(* IEC 61131-3 sources: RootPLC/conformance/cases/blocks, 22 files *)

(* ---- ok_rb_round4.st ---- *)
(* spec: [blocks.fault] [blocks.testable]
   expect: ok
   libraries: RootBlocks *)
(* Test suites of RB_SetpointProfile (F06.PROFILE), RB_Homing (F05.HOMING),
   RB_DataLog (F11.LOG), RB_ScaleOut (F01.SCALE.OUT) and RB_Drum
   (F05.DRUM). Every call passes the inputs that matter: block inputs keep
   their last value. *)
FUNCTION_BLOCK FB_Profile2
VAR_OUTPUT
    tg : ARRAY[1..8] OF REAL;
    rt : ARRAY[1..8] OF TIME;
    st : ARRAY[1..8] OF TIME;
END_VAR
tg[1] := 100.0; rt[1] := T#10s; st[1] := T#5s;
tg[2] := 50.0;  rt[2] := T#5s;  st[2] := T#2s;
END_FUNCTION_BLOCK

TEST profile_ramps_and_soaks
VAR p : RB_SetpointProfile; d : FB_Profile2; END_VAR
d();
p(PV := 20.0, Count := 2, Targets := d.tg, RampTimes := d.rt, SoakTimes := d.st);
ASSERT_FALSE(p.Busy);
ASSERT_EQ(0, p.Segment);
ADVANCE(T#1s);
p(Start := TRUE);
ASSERT_TRUE(p.Busy);
ASSERT_EQ(1, p.Segment);
ASSERT_TRUE(ABS(p.SP - 20.0) < 0.001);
ADVANCE(T#5s);
p(Start := FALSE);
ASSERT_TRUE(ABS(p.SP - 60.0) < 0.01);
ASSERT_FALSE(p.Soaking);
ADVANCE(T#5s);
p();
ASSERT_TRUE(ABS(p.SP - 100.0) < 0.001);
ASSERT_TRUE(p.Soaking);
ADVANCE(T#4900ms);
p();
ASSERT_EQ(1, p.Segment);
ADVANCE(T#100ms);
p();
ASSERT_EQ(2, p.Segment);
ASSERT_FALSE(p.Soaking);
ADVANCE(T#2500ms);
p();
ASSERT_TRUE(ABS(p.SP - 75.0) < 0.01);
ADVANCE(T#2500ms);
p();
ASSERT_TRUE(ABS(p.SP - 50.0) < 0.001);
ADVANCE(T#2s);
p();
ASSERT_TRUE(p.Done);
ASSERT_FALSE(p.Busy);
ASSERT_EQ(0, p.Segment);
ASSERT_TRUE(ABS(p.SP - 50.0) < 0.001);
(* a new start clears Done *)
p(Start := TRUE, PV := 30.0);
ASSERT_FALSE(p.Done);
ASSERT_TRUE(ABS(p.SP - 30.0) < 0.001);
END_TEST

TEST profile_hold_guarantee_and_abort
VAR p : RB_SetpointProfile; d : FB_Profile2; END_VAR
d();
p(PV := 20.0, Count := 1, Targets := d.tg, RampTimes := d.rt, SoakTimes := d.st, Start := TRUE);
ADVANCE(T#5s);
p(Start := FALSE);
ASSERT_TRUE(ABS(p.SP - 60.0) < 0.01);
ADVANCE(T#10s);
p(Hold := TRUE);
ASSERT_TRUE(ABS(p.SP - 60.0) < 0.01);
p(Hold := FALSE);
ADVANCE(T#5s);
p(Band := 2.0);
ASSERT_TRUE(p.Soaking);
(* guaranteed soak: PV far from SP, the soak waits *)
ADVANCE(T#10s);
p(PV := 90.0);
ASSERT_TRUE(p.Soaking);
ASSERT_EQ(1, p.Segment);
ADVANCE(T#1s);
p(PV := 98.0);
(* each call counts the time since the previous one *)
ADVANCE(T#3s);
p(PV := 98.0);
ASSERT_TRUE(p.Busy);
ADVANCE(T#1s);
p(PV := 98.0);
ASSERT_TRUE(p.Done);
(* abort while soaking *)
p(Start := TRUE, PV := 100.0);
ASSERT_TRUE(p.Busy);
ADVANCE(T#10s);
p(Start := FALSE);
ASSERT_TRUE(p.Soaking);
p(Abort := TRUE);
ASSERT_FALSE(p.Soaking);
ASSERT_FALSE(p.Busy);
ASSERT_EQ(0, p.Segment);
ASSERT_FALSE(p.Done);
ADVANCE(T#20s);
p(Abort := FALSE);
ASSERT_FALSE(p.Busy);
END_TEST

TEST profile_zero_times_and_count
VAR p : RB_SetpointProfile; tg : ARRAY[1..8] OF REAL; rt, st : ARRAY[1..8] OF TIME; END_VAR
tg[1] := 70.0;
p(PV := 10.0, Count := 0, Targets := tg, RampTimes := rt, SoakTimes := st, Start := TRUE);
ASSERT_TRUE(p.Error);
ASSERT_EQ(UDINT#1, p.ErrorID);
ASSERT_FALSE(p.Busy);
p(Start := FALSE, Count := 9);
p(Start := TRUE);
ASSERT_TRUE(p.Error);
p(Start := FALSE, Count := 8);
p(Start := TRUE);
ASSERT_FALSE(p.Error);
ASSERT_EQ(UDINT#0, p.ErrorID);
(* T#0s ramp and soak: a step to the target, one segment per call *)
p(Start := FALSE);
ASSERT_TRUE(ABS(p.SP - 70.0) < 0.001);
p();
ASSERT_EQ(2, p.Segment);
p(Count := 1);
p();
ASSERT_TRUE(p.Done);
(* a start with a bad count while running ends the program *)
p(Count := 8);
p(Start := TRUE);
p(Start := FALSE);
p();
ASSERT_EQ(2, p.Segment);
p(Count := 0);
p(Start := TRUE);
ASSERT_EQ(0, p.Segment);
ASSERT_FALSE(p.Busy);
END_TEST

TEST homing_seeks_and_backs_off
VAR h : RB_Homing; END_VAR
h();
ASSERT_FALSE(h.Busy OR h.Homed);
h(Start := TRUE);
ASSERT_TRUE(h.MoveToHome);
ASSERT_FALSE(h.MoveAway OR h.Slow);
ASSERT_TRUE(h.Busy);
ADVANCE(T#20s);
h(Start := FALSE, HomeSwitch := TRUE);
ASSERT_FALSE(h.MoveToHome);
ASSERT_TRUE(h.MoveAway AND h.Slow);
(* each phase has its own Timeout *)
ADVANCE(T#20s);
h();
ASSERT_FALSE(h.Error);
h(HomeSwitch := FALSE);
ASSERT_TRUE(h.Homed);
ASSERT_FALSE(h.Busy OR h.MoveAway OR h.MoveToHome);
(* starting on the switch: straight to backing off; Homed clears *)
h(Start := TRUE, HomeSwitch := TRUE);
ASSERT_FALSE(h.Homed);
ASSERT_TRUE(h.MoveAway);
h(Start := FALSE, HomeSwitch := FALSE);
ASSERT_TRUE(h.Homed);
(* a new start while seeking restarts the timing *)
h(Start := TRUE, Timeout := T#2s);
ADVANCE(T#1500ms);
h(Start := FALSE);
h(Start := TRUE);
ADVANCE(T#1500ms);
h(Start := FALSE);
ASSERT_FALSE(h.Error);
ASSERT_TRUE(h.MoveToHome);
h(Timeout := T#30s);
(* abort *)
h(Start := TRUE);
ASSERT_TRUE(h.MoveToHome);
h(Start := FALSE, Abort := TRUE);
ASSERT_FALSE(h.Busy OR h.MoveToHome OR h.Homed);
h(Start := TRUE);
ASSERT_FALSE(h.Busy);
END_TEST

TEST homing_timeouts
VAR h : RB_Homing; END_VAR
h(Start := TRUE, Timeout := T#2s);
ADVANCE(T#1900ms);
h();
ASSERT_FALSE(h.Error);
ADVANCE(T#100ms);
h();
ASSERT_TRUE(h.Error);
ASSERT_EQ(UDINT#1, h.ErrorID);
ASSERT_FALSE(h.MoveToHome OR h.Busy);
(* no start while the fault lasts *)
h(Start := FALSE);
h(Start := TRUE);
ASSERT_FALSE(h.Busy);
h(Start := FALSE, Reset := TRUE);
ASSERT_FALSE(h.Error);
ASSERT_EQ(UDINT#0, h.ErrorID);
h(Reset := FALSE, Start := TRUE);
ASSERT_TRUE(h.MoveToHome);
h(Start := FALSE, HomeSwitch := TRUE);
ADVANCE(T#2s);
h();
ASSERT_TRUE(h.Error);
ASSERT_EQ(UDINT#2, h.ErrorID);
ASSERT_FALSE(h.MoveAway OR h.Slow);
ASSERT_FALSE(h.Homed);
END_TEST

TEST data_log_ring_and_statistics
VAR l : RB_DataLog; i : INT; END_VAR
l(Value := 0.0, Enable := FALSE);
ASSERT_EQ(0, l.Count);
ASSERT_EQ(0, l.Newest);
l(Value := 5.0, Enable := TRUE);
ASSERT_EQ(1, l.Count);
ASSERT_EQ(1, l.Newest);
ASSERT_TRUE(ABS(l.Minimum - 5.0) < 0.001 AND ABS(l.Maximum - 5.0) < 0.001 AND ABS(l.Average - 5.0) < 0.001);
ADVANCE(T#500ms);
l(Value := 9.0);
ASSERT_EQ(1, l.Count);
ADVANCE(T#500ms);
l(Value := 1.0);
ASSERT_EQ(2, l.Count);
ASSERT_TRUE(ABS(l.Samples[2] - 1.0) < 0.001);
ASSERT_TRUE(ABS(l.Minimum - 1.0) < 0.001);
ASSERT_TRUE(ABS(l.Maximum - 5.0) < 0.001);
ASSERT_TRUE(ABS(l.Average - 3.0) < 0.001);
(* fill and wrap: 70 samples in all *)
FOR i := 3 TO 70 DO
    ADVANCE(T#1s);
    l(Value := INT_TO_REAL(i));
END_FOR;
ASSERT_EQ(64, l.Count);
ASSERT_EQ(6, l.Newest);
ASSERT_TRUE(ABS(l.Samples[6] - 70.0) < 0.001);
ASSERT_TRUE(ABS(l.Minimum - 7.0) < 0.001);
ASSERT_TRUE(ABS(l.Maximum - 70.0) < 0.001);
ASSERT_TRUE(ABS(l.Average - 38.5) < 0.001);
(* the next sample comes one Interval later, not before *)
ADVANCE(T#500ms);
l(Value := 71.0);
ASSERT_EQ(6, l.Newest);
ADVANCE(T#500ms);
l(Value := 71.0);
ASSERT_EQ(7, l.Newest);
(* paused, then cleared *)
ADVANCE(T#5s);
l(Value := 99.0, Enable := FALSE);
ASSERT_TRUE(ABS(l.Maximum - 71.0) < 0.001);
l(Clear := TRUE);
ASSERT_EQ(0, l.Count);
ASSERT_TRUE(ABS(l.Average) < 0.001 AND ABS(l.Maximum) < 0.001 AND ABS(l.Minimum) < 0.001);
l(Clear := FALSE, Enable := TRUE, Value := -4.0);
ASSERT_EQ(1, l.Newest);
ASSERT_TRUE(ABS(l.Minimum + 4.0) < 0.001 AND ABS(l.Maximum + 4.0) < 0.001);
END_TEST

TEST scale_out_to_an_output_word
VAR s : RB_ScaleOut; END_VAR
s(Value := 50.0);
ASSERT_EQ(13824, s.Raw);
ASSERT_FALSE(s.Limited OR s.Error);
s(Value := 100.0);
ASSERT_EQ(27648, s.Raw);
ASSERT_FALSE(s.Limited);
s(Value := 120.0);
ASSERT_EQ(27648, s.Raw);
ASSERT_TRUE(s.Limited);
s(Value := -5.0);
ASSERT_EQ(0, s.Raw);
ASSERT_TRUE(s.Limited);
s(Value := 0.5);
ASSERT_EQ(138, s.Raw);
s(Value := 0.0);
ASSERT_EQ(0, s.Raw);
ASSERT_FALSE(s.Limited);
(* the fail value on a fault *)
s(Value := 50.0, Fault := TRUE, FailValue := 25.0);
ASSERT_EQ(6912, s.Raw);
s(Fault := FALSE);
ASSERT_EQ(13824, s.Raw);
(* a reversed range and a live-zero raw range *)
s(Value := 25.0, EngMin := 100.0, EngMax := 0.0);
ASSERT_EQ(20736, s.Raw);
s(Value := 50.0, EngMin := 0.0, EngMax := 100.0, RawMin := 5530.0);
ASSERT_EQ(16589, s.Raw);
s(EngMax := 0.0);
ASSERT_TRUE(s.Error);
ASSERT_EQ(UDINT#1, s.ErrorID);
ASSERT_EQ(5530, s.Raw);
ASSERT_FALSE(s.Limited);
s(EngMax := 200.0);
ASSERT_FALSE(s.Error);
ASSERT_EQ(UDINT#0, s.ErrorID);
END_TEST

TEST drum_steps_by_time_and_event
VAR d : RB_Drum; p : ARRAY[1..16] OF WORD; t : ARRAY[1..16] OF TIME; END_VAR
p[1] := WORD#16#0001; p[2] := WORD#16#0006; p[3] := WORD#16#0010;
t[1] := T#2s; t[2] := T#0s; t[3] := T#1s;
d(Patterns := p, Times := t, Count := 3);
ASSERT_EQ(1, d.StepNo);
ASSERT_EQ(WORD#16#0001, d.Out);
ADVANCE(T#5s);
d();
ASSERT_EQ(1, d.StepNo);
d(Run := TRUE);
ADVANCE(T#1900ms);
d();
ASSERT_EQ(1, d.StepNo);
ASSERT_EQ(T#1900ms, d.StepTime);
ADVANCE(T#100ms);
d();
ASSERT_EQ(2, d.StepNo);
ASSERT_EQ(WORD#16#0006, d.Out);
ASSERT_EQ(T#0s, d.StepTime);
(* T#0s: waits for Next *)
ADVANCE(T#10s);
d();
ASSERT_EQ(2, d.StepNo);
d(Next := TRUE);
ASSERT_EQ(3, d.StepNo);
d(Next := FALSE);
(* paused while Run is FALSE *)
ADVANCE(T#500ms);
d();
ADVANCE(T#100ms);
d(Run := FALSE);
ADVANCE(T#100ms);
d(Run := FALSE);
ADVANCE(T#100ms);
d(Run := TRUE);
ADVANCE(T#300ms);
d();
ASSERT_EQ(3, d.StepNo);
ADVANCE(T#100ms);
d();
ASSERT_EQ(1, d.StepNo);
END_TEST

TEST drum_one_shot_reset_and_count
VAR d : RB_Drum; p : ARRAY[1..16] OF WORD; t : ARRAY[1..16] OF TIME; END_VAR
p[1] := WORD#16#00F0; p[2] := WORD#16#0F00;
d(Patterns := p, Times := t, Count := 2, Cyclic := FALSE);
d(Next := TRUE);
ASSERT_EQ(2, d.StepNo);
d(Next := FALSE);
d(Next := TRUE);
ASSERT_TRUE(d.Done);
ASSERT_EQ(2, d.StepNo);
ASSERT_EQ(WORD#16#0F00, d.Out);
d(Next := FALSE);
d(Next := TRUE);
ASSERT_EQ(2, d.StepNo);
d(Next := FALSE, Reset := TRUE);
ASSERT_EQ(1, d.StepNo);
ASSERT_FALSE(d.Done);
d(Reset := FALSE, Count := 0);
ASSERT_TRUE(d.Error);
ASSERT_EQ(UDINT#1, d.ErrorID);
ASSERT_EQ(WORD#0, d.Out);
ASSERT_EQ(0, d.StepNo);
d(Count := 17);
ASSERT_TRUE(d.Error);
d(Count := 1);
ASSERT_FALSE(d.Error);
ASSERT_EQ(1, d.StepNo);
d(Count := 16);
ASSERT_FALSE(d.Error);
ASSERT_EQ(UDINT#0, d.ErrorID);
ASSERT_EQ(1, d.StepNo);
(* a smaller Count while beyond it: back to step 1 *)
d(Next := TRUE);
d(Next := FALSE);
d(Next := TRUE);
d(Next := FALSE);
ASSERT_EQ(3, d.StepNo);
d(Count := 2);
ASSERT_EQ(1, d.StepNo);
END_TEST

(* ---- ok_rb_sequence.st ---- *)
(* spec: [blocks.command] [blocks.fault] [blocks.testable]
   expect: ok
   libraries: RootBlocks *)
(* Test suites of RB_StepChain (F05.STEPS) and RB_Phase (F05.PHASE). *)

(* the pattern the card shows: the chain, then the actions per step *)
FUNCTION_BLOCK FillCycle
VAR_INPUT
    start  : BOOL;
    full   : BOOL;
    empty  : BOOL;
END_VAR
VAR_OUTPUT
    inlet  : BOOL;
    outlet : BOOL;
    fills  : INT;
END_VAR
VAR
    chain : RB_StepChain;
END_VAR
CASE chain.StepNo OF
1: chain(Start := start, Proceed := full, LastStep := 2, StepTimeout := T#5s);
2: chain(Start := start, Proceed := empty, LastStep := 2, StepTimeout := T#5s);
ELSE
    chain(Start := start, Proceed := FALSE, LastStep := 2, StepTimeout := T#5s);
END_CASE;
inlet := chain.StepNo = 1;
outlet := chain.StepNo = 2;
IF chain.FirstCall AND chain.StepNo = 1 THEN
    fills := fills + 1;
END_IF;
END_FUNCTION_BLOCK

TEST chain_runs_its_steps_in_order
VAR f : FillCycle; END_VAR
f(start := FALSE);
ASSERT_EQ(0, f.chain.StepNo);
ASSERT_FALSE(f.chain.Busy);
f(start := TRUE);
ASSERT_EQ(1, f.chain.StepNo);
ASSERT_TRUE(f.inlet);
ASSERT_TRUE(f.chain.FirstCall);
ASSERT_TRUE(f.chain.Busy);
ASSERT_EQ(1, f.fills);
f(start := TRUE);
ASSERT_FALSE(f.chain.FirstCall);
ASSERT_EQ(1, f.fills);
f(start := TRUE, full := TRUE);
ASSERT_EQ(2, f.chain.StepNo);
ASSERT_TRUE(f.chain.FirstCall);
ASSERT_TRUE(f.outlet);
f(start := TRUE, full := TRUE, empty := TRUE);
ASSERT_EQ(0, f.chain.StepNo);
ASSERT_TRUE(f.chain.Done);
ASSERT_FALSE(f.chain.Busy);
f(start := TRUE, full := TRUE, empty := TRUE);
ASSERT_FALSE(f.chain.Done);
ASSERT_EQ(0, f.chain.StepNo);
(* a new rising edge starts it again *)
f(start := FALSE);
f(start := TRUE);
ASSERT_EQ(1, f.chain.StepNo);
ASSERT_EQ(2, f.fills);
END_TEST

TEST chain_step_time_and_timeout
VAR c : RB_StepChain; END_VAR
c(Start := TRUE, LastStep := 3, StepTimeout := T#2s);
ADVANCE(T#1500ms);
c(Start := TRUE, LastStep := 3, StepTimeout := T#2s);
ASSERT_TRUE(c.StepTime = T#1500ms);
ASSERT_FALSE(c.Error);
ADVANCE(T#500ms);
c(Start := TRUE, LastStep := 3, StepTimeout := T#2s);
ASSERT_TRUE(c.Error);
ASSERT_EQ(UDINT#1, c.ErrorID);
ASSERT_EQ(1, c.StepNo);
(* the fault holds the chain: Proceed is ignored *)
c(Start := TRUE, Proceed := TRUE, LastStep := 3, StepTimeout := T#2s);
ASSERT_EQ(1, c.StepNo);
(* reset restarts the step timer *)
c(Start := TRUE, Proceed := FALSE, LastStep := 3, StepTimeout := T#2s, Reset := TRUE);
ASSERT_FALSE(c.Error);
ASSERT_EQ(UDINT#0, c.ErrorID);
ASSERT_TRUE(c.StepTime = T#0s);
ADVANCE(T#1s);
c(Start := TRUE, Proceed := TRUE, LastStep := 3, StepTimeout := T#2s, Reset := FALSE);
ASSERT_EQ(2, c.StepNo);
ASSERT_TRUE(c.StepTime = T#0s);
(* no timeout configured: no fault *)
ADVANCE(T#1h);
c(Start := TRUE, Proceed := FALSE, LastStep := 3, StepTimeout := T#0s);
ASSERT_FALSE(c.Error);
END_TEST

TEST chain_hold_pauses_and_abort_resets
VAR c : RB_StepChain; END_VAR
c(Start := TRUE, LastStep := 2, StepTimeout := T#2s);
ADVANCE(T#1s);
c(Start := TRUE, Hold := TRUE, Proceed := TRUE, LastStep := 2, StepTimeout := T#2s);
ASSERT_EQ(1, c.StepNo);
ASSERT_TRUE(c.Held);
ADVANCE(T#10s);
c(Start := TRUE, Hold := TRUE, Proceed := FALSE, LastStep := 2, StepTimeout := T#2s);
ASSERT_FALSE(c.Error);
ASSERT_TRUE(c.StepTime = T#0s);
c(Start := TRUE, Hold := FALSE, Proceed := FALSE, LastStep := 2, StepTimeout := T#2s);
ASSERT_FALSE(c.Held);
ASSERT_FALSE(c.Error);
c(Start := TRUE, Abort := TRUE, LastStep := 2, StepTimeout := T#2s);
ASSERT_EQ(0, c.StepNo);
ASSERT_TRUE(c.Aborted);
ASSERT_FALSE(c.Busy);
ASSERT_FALSE(c.Held);
c(Start := TRUE, Abort := TRUE, LastStep := 2, StepTimeout := T#2s);
ASSERT_FALSE(c.Aborted);
(* while Abort is TRUE the chain does not start *)
c(Start := FALSE, Abort := TRUE, LastStep := 2);
c(Start := TRUE, Abort := TRUE, LastStep := 2);
ASSERT_EQ(0, c.StepNo);
END_TEST

TEST chain_branches_with_next_step
VAR c : RB_StepChain; END_VAR
c(Start := TRUE, LastStep := 5);
c(Start := TRUE, Proceed := TRUE, NextStep := 4, LastStep := 5);
ASSERT_EQ(4, c.StepNo);
ASSERT_TRUE(c.FirstCall);
c(Start := TRUE, Proceed := TRUE, NextStep := 0, LastStep := 5);
ASSERT_EQ(5, c.StepNo);
(* a jump back from the last step keeps the chain running *)
c(Start := TRUE, Proceed := TRUE, NextStep := 2, LastStep := 5);
ASSERT_EQ(2, c.StepNo);
ASSERT_FALSE(c.Done);
(* an abort with an active timeout fault clears it *)
c(Start := TRUE, Proceed := FALSE, StepTimeout := T#1s, LastStep := 5);
ADVANCE(T#2s);
c(Start := TRUE, Proceed := FALSE, StepTimeout := T#1s, LastStep := 5);
ASSERT_TRUE(c.Error);
c(Start := TRUE, Abort := TRUE, LastStep := 5);
ASSERT_FALSE(c.Error);
ASSERT_EQ(UDINT#0, c.ErrorID);
END_TEST

TEST phase_runs_holds_and_completes
VAR p : RB_Phase; END_VAR
p();
ASSERT_TRUE(p.State = RB_PHASE_STATE#Idle);
p(Start := TRUE);
ASSERT_TRUE(p.State = RB_PHASE_STATE#Running);
ASSERT_TRUE(p.Running);
ASSERT_FALSE(p.Rejected);
p(Start := FALSE, Hold := TRUE);
ASSERT_TRUE(p.State = RB_PHASE_STATE#Held);
ASSERT_FALSE(p.Running);
p(Hold := FALSE, Finished := TRUE);
ASSERT_TRUE(p.State = RB_PHASE_STATE#Held);
p(Restart := TRUE, Finished := FALSE);
ASSERT_TRUE(p.State = RB_PHASE_STATE#Running);
p(Restart := FALSE, Finished := TRUE);
ASSERT_TRUE(p.State = RB_PHASE_STATE#Complete);
ASSERT_TRUE(p.Done);
p(Finished := FALSE, Reset := TRUE);
ASSERT_TRUE(p.State = RB_PHASE_STATE#Idle);
ASSERT_FALSE(p.Done);
END_TEST

TEST phase_stop_abort_and_rejected_commands
VAR p : RB_Phase; END_VAR
(* commands that do not fit the state are rejected *)
p(Hold := TRUE);
ASSERT_TRUE(p.Rejected);
ASSERT_TRUE(p.State = RB_PHASE_STATE#Idle);
p(Hold := FALSE, Restart := TRUE);
ASSERT_TRUE(p.Rejected);
p(Restart := FALSE, Stop := TRUE);
ASSERT_TRUE(p.Rejected);
p(Stop := FALSE, Abort := TRUE);
ASSERT_TRUE(p.Rejected);
p(Abort := FALSE, Reset := TRUE);
ASSERT_TRUE(p.Rejected);
p(Reset := FALSE);
ASSERT_FALSE(p.Rejected);
p(Start := TRUE);
ASSERT_FALSE(p.Rejected);
p(Start := FALSE);
p(Start := TRUE);
ASSERT_TRUE(p.Rejected);
ASSERT_TRUE(p.State = RB_PHASE_STATE#Running);
(* stop from running, abort from stopped, reset from aborted *)
p(Start := FALSE, Stop := TRUE);
ASSERT_TRUE(p.State = RB_PHASE_STATE#Stopped);
p(Stop := FALSE, Abort := TRUE);
ASSERT_TRUE(p.State = RB_PHASE_STATE#Aborted);
p(Abort := FALSE, Stop := TRUE);
ASSERT_TRUE(p.Rejected);
p(Stop := FALSE, Reset := TRUE);
ASSERT_TRUE(p.State = RB_PHASE_STATE#Idle);
(* stop and abort from held; reset from stopped *)
p(Reset := FALSE, Start := TRUE);
p(Start := FALSE, Hold := TRUE);
p(Hold := FALSE, Stop := TRUE);
ASSERT_TRUE(p.State = RB_PHASE_STATE#Stopped);
p(Stop := FALSE, Reset := TRUE);
ASSERT_TRUE(p.State = RB_PHASE_STATE#Idle);
p(Reset := FALSE, Start := TRUE);
p(Start := FALSE, Hold := TRUE);
p(Hold := FALSE, Abort := TRUE);
ASSERT_TRUE(p.State = RB_PHASE_STATE#Aborted);
(* abort from running; completed phases reject stop *)
p(Abort := FALSE, Reset := TRUE);
p(Reset := FALSE, Start := TRUE);
p(Start := FALSE, Abort := TRUE);
ASSERT_TRUE(p.State = RB_PHASE_STATE#Aborted);
p(Abort := FALSE, Reset := TRUE);
p(Reset := FALSE, Start := TRUE);
p(Start := FALSE, Finished := TRUE);
p(Finished := FALSE, Stop := TRUE);
ASSERT_TRUE(p.Rejected);
ASSERT_TRUE(p.State = RB_PHASE_STATE#Complete);
p(Stop := FALSE, Abort := TRUE);
ASSERT_TRUE(p.Rejected);
p(Abort := FALSE, Hold := TRUE);
ASSERT_TRUE(p.Rejected);
END_TEST

TEST phase_highest_valid_command_acts
VAR p : RB_Phase; END_VAR
(* in idle an abort is invalid: the start given with it acts, and the
   abort is reported as rejected *)
p(Start := TRUE, Abort := TRUE);
ASSERT_TRUE(p.State = RB_PHASE_STATE#Running);
ASSERT_TRUE(p.Rejected);
(* running: abort and hold together, abort wins; the hold was valid, so
   nothing is rejected *)
p(Start := FALSE, Abort := FALSE);
p(Abort := TRUE, Hold := TRUE);
ASSERT_TRUE(p.State = RB_PHASE_STATE#Aborted);
ASSERT_FALSE(p.Rejected);
(* aborted: reset and start together; start is invalid there, reset acts *)
p(Abort := FALSE, Hold := FALSE);
p(Reset := TRUE, Start := TRUE);
ASSERT_TRUE(p.State = RB_PHASE_STATE#Idle);
ASSERT_TRUE(p.Rejected);
(* idle: a restart (invalid) and a start: start acts *)
p(Reset := FALSE, Start := FALSE);
p(Restart := TRUE, Start := TRUE);
ASSERT_TRUE(p.State = RB_PHASE_STATE#Running);
ASSERT_TRUE(p.Rejected);
(* running: a command acting keeps Finished from completing in that call *)
p(Restart := FALSE, Start := FALSE);
p(Hold := TRUE, Finished := TRUE);
ASSERT_TRUE(p.State = RB_PHASE_STATE#Held);
(* held: stop and restart together; stop wins, restart was valid *)
p(Hold := FALSE, Finished := FALSE);
p(Stop := TRUE, Restart := TRUE);
ASSERT_TRUE(p.State = RB_PHASE_STATE#Stopped);
ASSERT_FALSE(p.Rejected);
(* stopped: a stop again is invalid *)
p(Stop := FALSE, Restart := FALSE);
p(Stop := TRUE);
ASSERT_TRUE(p.Rejected);
ASSERT_TRUE(p.State = RB_PHASE_STATE#Stopped);
END_TEST

(* ---- ok_rb_alarm.st ---- *)
(* spec: [blocks.testable] [blocks.library]
   expect: ok
   libraries: RootBlocks *)
(* Test suite of RB_Alarm (F08.ALARM). Every call passes the inputs that
   matter: block inputs keep their last value. *)
TEST alarm_states_with_acknowledge_while_active
VAR a : RB_Alarm; END_VAR
a(In := FALSE);
ASSERT_TRUE(a.State = RB_ALARM_STATE#Normal);
a(In := TRUE);
ASSERT_TRUE(a.Active);
ASSERT_TRUE(a.Unacked);
ASSERT_TRUE(a.State = RB_ALARM_STATE#ActiveUnack);
ASSERT_EQ(UDINT#1, a.Count);
a(In := TRUE, Ack := TRUE);
ASSERT_FALSE(a.Unacked);
ASSERT_TRUE(a.State = RB_ALARM_STATE#ActiveAcked);
a(In := TRUE, Ack := FALSE);
ASSERT_EQ(UDINT#1, a.Count);
a(In := FALSE);
ASSERT_FALSE(a.Active);
ASSERT_TRUE(a.State = RB_ALARM_STATE#Normal);
END_TEST

TEST alarm_returns_unacknowledged
VAR a : RB_Alarm; END_VAR
a(In := TRUE);
a(In := FALSE);
ASSERT_FALSE(a.Active);
ASSERT_TRUE(a.Unacked);
ASSERT_TRUE(a.State = RB_ALARM_STATE#ReturnedUnack);
a(In := FALSE, Ack := TRUE);
ASSERT_TRUE(a.State = RB_ALARM_STATE#Normal);
a(In := TRUE, Ack := TRUE);
ASSERT_TRUE(a.State = RB_ALARM_STATE#ActiveUnack);
ASSERT_EQ(UDINT#2, a.Count);
END_TEST

TEST alarm_delays
VAR a : RB_Alarm; END_VAR
a(In := TRUE, OnDelay := T#2s, OffDelay := T#1s);
ASSERT_FALSE(a.Active);
ADVANCE(T#1900ms);
a(In := TRUE, OnDelay := T#2s, OffDelay := T#1s);
ASSERT_FALSE(a.Active);
ADVANCE(T#200ms);
a(In := TRUE, OnDelay := T#2s, OffDelay := T#1s);
ASSERT_TRUE(a.Active);
a(In := FALSE, OnDelay := T#2s, OffDelay := T#1s);
ADVANCE(T#900ms);
a(In := FALSE, OnDelay := T#2s, OffDelay := T#1s);
ASSERT_TRUE(a.Active);
ADVANCE(T#200ms);
a(In := FALSE, OnDelay := T#2s, OffDelay := T#1s);
ASSERT_FALSE(a.Active);
ASSERT_TRUE(a.State = RB_ALARM_STATE#ReturnedUnack);
END_TEST

TEST alarm_out_of_service
VAR a : RB_Alarm; END_VAR
a(In := TRUE);
a(In := TRUE, Enable := FALSE);
ASSERT_FALSE(a.Active);
ASSERT_FALSE(a.Unacked);
ASSERT_TRUE(a.State = RB_ALARM_STATE#Normal);
a(In := TRUE, Enable := FALSE);
ASSERT_EQ(UDINT#1, a.Count);
a(In := TRUE, Enable := TRUE);
ASSERT_TRUE(a.Active);
ASSERT_EQ(UDINT#2, a.Count);
END_TEST

(* ---- ok_rb_control.st ---- *)
(* spec: [blocks.mode] [blocks.fault] [blocks.testable]
   expect: ok
   libraries: RootBlocks *)
(* Test suites of RB_PID (F06.PID) and RB_OnOff (F06.ONOFF). Every call
   passes the inputs that matter: block inputs keep their last value. *)
TEST pid_proportional_both_actions
VAR c : RB_PID; d : RB_PID; END_VAR
c(Mode := RB_MODE#Auto, SP := 50.0, PV := 40.0, Kp := 2.0);
ASSERT_TRUE(ABS(c.Out - 20.0) < 0.001);
ASSERT_FALSE(c.Saturated);
d(Mode := RB_MODE#Auto, SP := 50.0, PV := 60.0, Kp := 2.0, Direct := TRUE);
ASSERT_TRUE(ABS(d.Out - 20.0) < 0.001);
d(Mode := RB_MODE#Auto, SP := 50.0, PV := 40.0, Kp := 2.0, Direct := TRUE);
ASSERT_TRUE(ABS(d.Out) < 0.001);
ASSERT_TRUE(d.Saturated);
END_TEST

TEST pid_integral_adds_up_over_time
VAR c : RB_PID; i : INT; END_VAR
c(Mode := RB_MODE#Auto, SP := 50.0, PV := 40.0, Kp := 1.0, Ti := T#1s);
ASSERT_TRUE(ABS(c.Out - 10.0) < 0.001);
FOR i := 1 TO 10 DO
    ADVANCE(T#100ms);
    c(Mode := RB_MODE#Auto, SP := 50.0, PV := 40.0, Kp := 1.0, Ti := T#1s);
END_FOR;
ASSERT_TRUE(ABS(c.Out - 20.0) < 0.001);
(* without integral time the output stays at the proportional part *)
ADVANCE(T#1s);
c(Mode := RB_MODE#Auto, SP := 50.0, PV := 40.0, Kp := 1.0, Ti := T#0s);
ASSERT_TRUE(ABS(c.Out - 10.0) < 0.001);
END_TEST

TEST pid_anti_windup_leaves_saturation_at_once
VAR c : RB_PID; i : INT; END_VAR
FOR i := 1 TO 100 DO
    ADVANCE(T#100ms);
    c(Mode := RB_MODE#Auto, SP := 60.0, PV := 0.0, Kp := 1.0, Ti := T#1s);
END_FOR;
ASSERT_TRUE(ABS(c.Out - 100.0) < 0.001);
ASSERT_TRUE(c.Saturated);
(* the error turns negative: the output leaves the limit in the same call *)
ADVANCE(T#100ms);
c(Mode := RB_MODE#Auto, SP := 60.0, PV := 61.0, Kp := 1.0, Ti := T#1s);
ASSERT_TRUE(c.Out < 100.0);
ASSERT_FALSE(c.Saturated);
(* and at the lower limit too *)
FOR i := 1 TO 100 DO
    ADVANCE(T#100ms);
    c(Mode := RB_MODE#Auto, SP := 0.0, PV := 60.0, Kp := 1.0, Ti := T#1s);
END_FOR;
ASSERT_TRUE(ABS(c.Out) < 0.001);
ADVANCE(T#100ms);
c(Mode := RB_MODE#Auto, SP := 61.0, PV := 60.0, Kp := 1.0, Ti := T#1s);
ASSERT_TRUE(c.Out > 0.0);
END_TEST

TEST pid_derivative_on_the_measurement
VAR c : RB_PID; d : RB_PID; END_VAR
c(Mode := RB_MODE#Auto, SP := 50.0, PV := 40.0, Kp := 1.0, Td := T#1s);
ASSERT_TRUE(ABS(c.Out - 10.0) < 0.001);
ADVANCE(T#100ms);
(* a set-point step: no derivative kick *)
c(Mode := RB_MODE#Auto, SP := 60.0, PV := 40.0, Kp := 1.0, Td := T#1s);
ASSERT_TRUE(ABS(c.Out - 20.0) < 0.001);
ADVANCE(T#100ms);
(* the measurement rises 1 in 0.1 s: D = -1 * 1 s * 10/s *)
c(Mode := RB_MODE#Auto, SP := 60.0, PV := 41.0, Kp := 1.0, Td := T#1s);
ASSERT_TRUE(ABS(c.Out - 9.0) < 0.001);
(* direct action: the sign of the derivative follows *)
d(Mode := RB_MODE#Auto, SP := 20.0, PV := 40.0, Kp := 1.0, Td := T#1s, Direct := TRUE);
ADVANCE(T#100ms);
d(Mode := RB_MODE#Auto, SP := 20.0, PV := 41.0, Kp := 1.0, Td := T#1s, Direct := TRUE);
ASSERT_TRUE(ABS(d.Out - 31.0) < 0.001);
(* two calls at the same instant: no derivative *)
d(Mode := RB_MODE#Auto, SP := 20.0, PV := 45.0, Kp := 1.0, Td := T#1s, Direct := TRUE);
ASSERT_TRUE(ABS(d.Out - 25.0) < 0.001);
END_TEST

TEST pid_manual_off_and_bumpless_transfer
VAR c : RB_PID; END_VAR
c(Mode := RB_MODE#Manual, SP := 50.0, PV := 50.0, Kp := 1.0, Ti := T#10s, ManValue := 40.0);
ASSERT_TRUE(ABS(c.Out - 40.0) < 0.001);
ASSERT_FALSE(c.Saturated);
c(Mode := RB_MODE#Manual, SP := 50.0, PV := 50.0, Kp := 1.0, Ti := T#10s, ManValue := 140.0);
ASSERT_TRUE(ABS(c.Out - 100.0) < 0.001);
ASSERT_FALSE(c.Saturated);
c(Mode := RB_MODE#Manual, SP := 50.0, PV := 50.0, Kp := 1.0, Ti := T#10s, ManValue := 40.0);
ADVANCE(T#100ms);
c(Mode := RB_MODE#Auto, SP := 50.0, PV := 50.0, Kp := 1.0, Ti := T#10s);
ASSERT_TRUE(ABS(c.Out - 40.0) < 0.001);
c(Mode := RB_MODE#Off, SP := 50.0, PV := 50.0, Kp := 1.0, Ti := T#10s, OutMin := 5.0);
ASSERT_TRUE(ABS(c.Out - 5.0) < 0.001);
ASSERT_FALSE(c.Saturated);
(* from Off, Auto starts at the minimum, not with a jump *)
ADVANCE(T#100ms);
c(Mode := RB_MODE#Auto, SP := 50.0, PV := 50.0, Kp := 1.0, Ti := T#10s, OutMin := 5.0);
ASSERT_TRUE(ABS(c.Out - 5.0) < 0.001);
ASSERT_TRUE(c.Saturated);
END_TEST

TEST pid_invalid_range_is_a_fault
VAR c : RB_PID; END_VAR
c(Mode := RB_MODE#Auto, SP := 50.0, PV := 40.0, Kp := 1.0, OutMin := 10.0, OutMax := 10.0);
ASSERT_TRUE(c.Error);
ASSERT_EQ(UDINT#1, c.ErrorID);
ASSERT_TRUE(ABS(c.Out - 10.0) < 0.001);
ASSERT_FALSE(c.Saturated);
c(Mode := RB_MODE#Auto, SP := 50.0, PV := 40.0, Kp := 1.0, OutMin := 0.0, OutMax := 100.0);
ASSERT_TRUE(c.Error);
c(Mode := RB_MODE#Auto, SP := 50.0, PV := 40.0, Kp := 1.0, OutMin := 0.0, OutMax := 100.0, Reset := TRUE);
ASSERT_FALSE(c.Error);
ASSERT_EQ(UDINT#0, c.ErrorID);
ASSERT_TRUE(ABS(c.Out - 10.0) < 0.001);
END_TEST

TEST onoff_heating_with_hysteresis
VAR h : RB_OnOff; END_VAR
h(Enable := TRUE, SP := 20.0, PV := 19.5, Hysteresis := 2.0);
ASSERT_FALSE(h.Out);
h(Enable := TRUE, SP := 20.0, PV := 19.0, Hysteresis := 2.0);
ASSERT_TRUE(h.Out);
h(Enable := TRUE, SP := 20.0, PV := 20.9, Hysteresis := 2.0);
ASSERT_TRUE(h.Out);
h(Enable := TRUE, SP := 20.0, PV := 21.0, Hysteresis := 2.0);
ASSERT_FALSE(h.Out);
h(Enable := TRUE, SP := 20.0, PV := 19.1, Hysteresis := 2.0);
ASSERT_FALSE(h.Out);
h(Enable := TRUE, SP := 20.0, PV := 18.0, Hysteresis := -2.0);
ASSERT_TRUE(h.Out);
h(Enable := FALSE, SP := 20.0, PV := 18.0, Hysteresis := 2.0);
ASSERT_FALSE(h.Out);
END_TEST

TEST onoff_cooling_with_hysteresis
VAR c : RB_OnOff; END_VAR
c(Enable := TRUE, SP := 5.0, PV := 6.0, Hysteresis := 2.0, Direct := TRUE);
ASSERT_TRUE(c.Out);
c(Enable := TRUE, SP := 5.0, PV := 4.1, Hysteresis := 2.0, Direct := TRUE);
ASSERT_TRUE(c.Out);
c(Enable := TRUE, SP := 5.0, PV := 4.0, Hysteresis := 2.0, Direct := TRUE);
ASSERT_FALSE(c.Out);
c(Enable := TRUE, SP := 5.0, PV := 5.9, Hysteresis := 2.0, Direct := TRUE);
ASSERT_FALSE(c.Out);
END_TEST

TEST pid_anti_windup_bounds_exactly
VAR c : RB_PID; i : INT; END_VAR
(* high limit: P = 60, the integral held at 40 *)
FOR i := 1 TO 50 DO
    ADVANCE(T#100ms);
    c(Mode := RB_MODE#Auto, SP := 60.0, PV := 0.0, Kp := 1.0, Ti := T#1s, Td := T#1s);
END_FOR;
(* the measurement rises 1 in 0.1 s: P = 59, D = -10, I = 40 + 5.9 *)
ADVANCE(T#100ms);
c(Mode := RB_MODE#Auto, SP := 60.0, PV := 1.0, Kp := 1.0, Ti := T#1s, Td := T#1s);
ASSERT_TRUE(ABS(c.Out - 94.9) < 0.01);
(* the error turns: P = -1, I = 45.9 - 0.1, D = 0 *)
ADVANCE(T#100ms);
c(Mode := RB_MODE#Auto, SP := 0.0, PV := 1.0, Kp := 1.0, Ti := T#1s, Td := T#1s);
ASSERT_TRUE(ABS(c.Out - 44.8) < 0.01);
(* low limit: P = -60 already holds the output at 0, so the integral
   (45.8) does not move further down and is not raised to cancel P *)
FOR i := 1 TO 50 DO
    ADVANCE(T#100ms);
    c(Mode := RB_MODE#Auto, SP := 0.0, PV := 60.0, Kp := 1.0, Ti := T#1s, Td := T#1s);
END_FOR;
ASSERT_TRUE(ABS(c.Out) < 0.01);
(* the measurement falls 1 in 0.1 s: P = -59, D = +10, I = 45.8: still 0 *)
ADVANCE(T#100ms);
c(Mode := RB_MODE#Auto, SP := 0.0, PV := 59.0, Kp := 1.0, Ti := T#1s, Td := T#1s);
ASSERT_TRUE(ABS(c.Out) < 0.01);
(* the error turns positive: P = 1, I = 45.8: the output follows gently *)
ADVANCE(T#100ms);
c(Mode := RB_MODE#Auto, SP := 60.0, PV := 59.0, Kp := 1.0, Ti := T#1s, Td := T#0s);
ASSERT_TRUE(ABS(c.Out - 46.9) < 0.01);
END_TEST

TEST pid_no_jump_after_a_long_saturation
VAR c : RB_PID; i : INT; END_VAR
(* pinned at the lower limit by a large error for 5 s *)
FOR i := 1 TO 50 DO
    ADVANCE(T#100ms);
    c(Mode := RB_MODE#Auto, SP := 0.0, PV := 73.6, Kp := 2.0, Ti := T#10s);
END_FOR;
ASSERT_TRUE(ABS(c.Out) < 0.001);
(* a small positive error gives a small output, not the upper limit *)
ADVANCE(T#100ms);
c(Mode := RB_MODE#Auto, SP := 75.0, PV := 73.6, Kp := 2.0, Ti := T#10s);
ASSERT_TRUE(c.Out > 2.0 AND c.Out < 3.5);
END_TEST

TEST pid_bumpless_with_an_error_present
VAR c : RB_PID; END_VAR
c(Mode := RB_MODE#Manual, SP := 50.0, PV := 45.0, Kp := 1.0, Ti := T#10s, ManValue := 40.0);
ADVANCE(T#100ms);
c(Mode := RB_MODE#Auto, SP := 50.0, PV := 45.0, Kp := 1.0, Ti := T#10s);
ASSERT_TRUE(ABS(c.Out - 40.05) < 0.001);
END_TEST

(* ---- ok_rb_control2.st ---- *)
(* spec: [blocks.fault] [blocks.testable]
   expect: ok
   libraries: RootBlocks *)
(* Test suites of RB_SplitRange (F06.SPLIT) and RB_AlarmSummary
   (F08.ALARM.SUMMARY). Every call passes the inputs that matter: block
   inputs keep their last value. *)
TEST split_range_sequential
VAR s : RB_SplitRange; END_VAR
s(In := 0.0);
ASSERT_TRUE(ABS(s.OutA) < 0.001 AND ABS(s.OutB) < 0.001);
ASSERT_FALSE(s.Error);
s(In := 25.0);
ASSERT_TRUE(ABS(s.OutA - 50.0) < 0.001);
ASSERT_TRUE(ABS(s.OutB) < 0.001);
s(In := 50.0);
ASSERT_TRUE(ABS(s.OutA - 100.0) < 0.001);
ASSERT_TRUE(ABS(s.OutB) < 0.001);
s(In := 75.0);
ASSERT_TRUE(ABS(s.OutA - 100.0) < 0.001);
ASSERT_TRUE(ABS(s.OutB - 50.0) < 0.001);
s(In := 100.0);
ASSERT_TRUE(ABS(s.OutB - 100.0) < 0.001);
s(In := 120.0);
ASSERT_TRUE(ABS(s.OutB - 100.0) < 0.001);
s(In := -10.0);
ASSERT_TRUE(ABS(s.OutA) < 0.001);
(* another split point *)
s(In := 30.0, SplitPoint := 60.0);
ASSERT_TRUE(ABS(s.OutA - 50.0) < 0.001);
s(In := 80.0);
ASSERT_TRUE(ABS(s.OutB - 50.0) < 0.001);
END_TEST

TEST split_range_heating_and_cooling
VAR s : RB_SplitRange; END_VAR
(* A cools below the split, B heats above it *)
s(In := 0.0, InvertA := TRUE);
ASSERT_TRUE(ABS(s.OutA - 100.0) < 0.001);
s(In := 25.0);
ASSERT_TRUE(ABS(s.OutA - 50.0) < 0.001);
s(In := 50.0);
ASSERT_TRUE(ABS(s.OutA) < 0.001);
ASSERT_TRUE(ABS(s.OutB) < 0.001);
s(In := 90.0);
ASSERT_TRUE(ABS(s.OutA) < 0.001);
ASSERT_TRUE(ABS(s.OutB - 80.0) < 0.001);
s(In := -10.0);
ASSERT_TRUE(ABS(s.OutA - 100.0) < 0.001);
END_TEST

TEST split_range_deadband
VAR s : RB_SplitRange; END_VAR
(* dead band 10: A over 0 .. 45, B over 55 .. 100 *)
s(In := 22.5, Deadband := 10.0);
ASSERT_TRUE(ABS(s.OutA - 50.0) < 0.001);
s(In := 50.0);
ASSERT_TRUE(ABS(s.OutA - 100.0) < 0.001);
ASSERT_TRUE(ABS(s.OutB) < 0.001);
s(In := 55.0);
ASSERT_TRUE(ABS(s.OutB) < 0.001);
s(In := 77.5);
ASSERT_TRUE(ABS(s.OutB - 50.0) < 0.001);
s(In := 22.5, InvertA := TRUE);
ASSERT_TRUE(ABS(s.OutA - 50.0) < 0.001);
END_TEST

TEST split_range_bad_settings
VAR s : RB_SplitRange; END_VAR
s(In := 75.0, SplitPoint := 0.0);
ASSERT_TRUE(s.Error);
ASSERT_EQ(UDINT#1, s.ErrorID);
ASSERT_TRUE(ABS(s.OutA) < 0.001 AND ABS(s.OutB) < 0.001);
s(SplitPoint := 100.0);
ASSERT_TRUE(s.Error);
s(SplitPoint := 95.0, Deadband := 10.0);
ASSERT_TRUE(s.Error);
s(SplitPoint := 5.0, Deadband := 10.0);
ASSERT_TRUE(s.Error);
s(SplitPoint := 50.0, Deadband := 10.0);
ASSERT_FALSE(s.Error);
ASSERT_EQ(UDINT#0, s.ErrorID);
s(SplitPoint := 1.0, Deadband := 0.0, In := 50.5);
ASSERT_FALSE(s.Error);
ASSERT_TRUE(ABS(s.OutB - 50.0) < 0.001);
s(SplitPoint := 99.0, In := 49.5);
ASSERT_FALSE(s.Error);
ASSERT_TRUE(ABS(s.OutA - 50.0) < 0.001);
END_TEST

TEST alarm_summary_counts_horn_and_first_out
VAR a : RB_AlarmSummary; st : ARRAY[1..32] OF RB_ALARM_STATE; END_VAR
a(States := st);
ASSERT_EQ(0, a.Active);
ASSERT_EQ(0, a.Unacked);
ASSERT_FALSE(a.Lamp OR a.Horn);
ASSERT_EQ(0, a.FirstOut);
st[5] := RB_ALARM_STATE#ActiveUnack;
a(States := st);
ASSERT_EQ(1, a.Active);
ASSERT_EQ(1, a.Unacked);
ASSERT_TRUE(a.Horn);
ASSERT_EQ(5, a.FirstOut);
(* silenced, then a second alarm sounds the horn again *)
a(States := st, Silence := TRUE);
ASSERT_FALSE(a.Horn);
a(States := st, Silence := FALSE);
ASSERT_FALSE(a.Horn);
st[3] := RB_ALARM_STATE#ActiveUnack;
a(States := st);
ASSERT_TRUE(a.Horn);
ASSERT_EQ(2, a.Active);
ASSERT_EQ(5, a.FirstOut);
(* both acknowledged: the horn stops, the lamp is steady *)
st[3] := RB_ALARM_STATE#ActiveAcked;
st[5] := RB_ALARM_STATE#ActiveAcked;
a(States := st);
ASSERT_FALSE(a.Horn);
ASSERT_EQ(0, a.Unacked);
ASSERT_EQ(2, a.Active);
ASSERT_TRUE(a.Lamp);
ADVANCE(T#600ms);
a(States := st);
ASSERT_TRUE(a.Lamp);
(* one returns unacknowledged: not active, but unacknowledged *)
st[5] := RB_ALARM_STATE#ReturnedUnack;
st[3] := RB_ALARM_STATE#Normal;
a(States := st);
ASSERT_EQ(0, a.Active);
ASSERT_EQ(1, a.Unacked);
ASSERT_EQ(5, a.FirstOut);
ASSERT_TRUE(a.Horn);
st[5] := RB_ALARM_STATE#Normal;
a(States := st);
ASSERT_EQ(0, a.FirstOut);
ASSERT_FALSE(a.Lamp OR a.Horn);
(* the next first-out is the lowest number active in one call *)
st[9] := RB_ALARM_STATE#ActiveAcked;
st[7] := RB_ALARM_STATE#ActiveUnack;
a(States := st);
ASSERT_EQ(7, a.FirstOut);
END_TEST

TEST alarm_summary_flashing_lamp
VAR a : RB_AlarmSummary; st : ARRAY[1..32] OF RB_ALARM_STATE; END_VAR
st[1] := RB_ALARM_STATE#ActiveUnack;
a(States := st);
ASSERT_TRUE(a.Lamp);
ADVANCE(T#400ms);
a(States := st);
ASSERT_TRUE(a.Lamp);
ADVANCE(T#100ms);
a(States := st);
ASSERT_FALSE(a.Lamp);
ADVANCE(T#500ms);
a(States := st);
ASSERT_TRUE(a.Lamp);
ADVANCE(T#500ms);
a(States := st);
ASSERT_FALSE(a.Lamp);
(* the timer restarts at each toggle *)
ADVANCE(T#100ms);
a(States := st);
ASSERT_FALSE(a.Lamp);
(* another rate *)
ADVANCE(T#100ms);
a(States := st, Blink := T#200ms);
ASSERT_TRUE(a.Lamp);
(* cleared while dark: the next alarm starts lit, with a full phase *)
ADVANCE(T#200ms);
a(States := st);
ASSERT_FALSE(a.Lamp);
st[1] := RB_ALARM_STATE#Normal;
a(States := st, Blink := T#500ms);
ASSERT_FALSE(a.Lamp);
ADVANCE(T#300ms);
a(States := st);
st[1] := RB_ALARM_STATE#ActiveUnack;
a(States := st);
ASSERT_TRUE(a.Lamp);
ADVANCE(T#400ms);
a(States := st);
ASSERT_TRUE(a.Lamp);
(* one acknowledged alarm: steady *)
st[1] := RB_ALARM_STATE#ActiveAcked;
a(States := st);
ASSERT_TRUE(a.Lamp);
END_TEST

TEST alarm_summary_unused_alarms
VAR a : RB_AlarmSummary; st : ARRAY[1..32] OF RB_ALARM_STATE; END_VAR
st[32] := RB_ALARM_STATE#ActiveUnack;
st[1] := RB_ALARM_STATE#ActiveUnack;
a(States := st, Used := DWORD#16#7FFFFFFE);
ASSERT_EQ(0, a.Active);
ASSERT_EQ(0, a.Unacked);
ASSERT_FALSE(a.Horn);
a(States := st, Used := DWORD#16#80000000);
ASSERT_EQ(1, a.Active);
ASSERT_EQ(32, a.FirstOut);
END_TEST

(* ---- ok_rb_cylinder.st ---- *)
(* spec: [blocks.command] [blocks.mode] [blocks.interlock] [blocks.fault] [blocks.feedback] [blocks.status]
   expect: ok
   libraries: RootBlocks *)
(* Test suite of RB_Cylinder (card blocks/cards/F04.CYLINDER.md). Every call
   passes the inputs that matter: block inputs keep their last value. *)
TEST cylinder_double_acting_strokes
VAR c : RB_Cylinder; END_VAR
c(Mode := RB_MODE#Auto, AutoExtend := FALSE, FbExtended := FALSE, FbRetracted := TRUE);
ASSERT_FALSE(c.Extend);
ASSERT_TRUE(c.Retract);
ASSERT_TRUE(c.IsRetracted);
c(Mode := RB_MODE#Auto, AutoExtend := TRUE, FbExtended := FALSE, FbRetracted := TRUE);
ASSERT_TRUE(c.Extend);
ASSERT_FALSE(c.Retract);
ASSERT_TRUE(c.Status.Commanded);
c(Mode := RB_MODE#Auto, AutoExtend := TRUE, FbExtended := TRUE, FbRetracted := FALSE);
ASSERT_TRUE(c.IsExtended);
ASSERT_FALSE(c.IsRetracted);
ASSERT_TRUE(c.Status.Active);
ASSERT_EQ(UDINT#1, c.Status.Starts);
ASSERT_TRUE(c.Status.Mode = RB_MODE#Auto);
c(Mode := RB_MODE#Auto, AutoExtend := TRUE, FbExtended := TRUE, FbRetracted := FALSE);
ASSERT_EQ(UDINT#1, c.Status.Starts);
ADVANCE(T#5s);
c(Mode := RB_MODE#Auto, AutoExtend := TRUE, FbExtended := TRUE, FbRetracted := FALSE);
ASSERT_FALSE(c.Error);
ASSERT_FALSE(c.Status.Error);
END_TEST

TEST cylinder_modes_interlock_permissive
VAR c : RB_Cylinder; END_VAR
c(Mode := RB_MODE#Auto, ManExtend := TRUE, FbRetracted := TRUE);
ASSERT_FALSE(c.Extend);
c(Mode := RB_MODE#Manual, ManExtend := TRUE, AutoExtend := FALSE, FbRetracted := TRUE);
ASSERT_TRUE(c.Extend);
c(Mode := RB_MODE#Manual, ManExtend := TRUE, Interlock := TRUE, FbRetracted := TRUE);
ASSERT_FALSE(c.Extend);
ASSERT_FALSE(c.Retract);
c(Mode := RB_MODE#Off, ManExtend := TRUE, AutoExtend := TRUE, Interlock := FALSE, FbRetracted := TRUE);
ASSERT_FALSE(c.Extend);
ASSERT_FALSE(c.Retract);
c(Mode := RB_MODE#Auto, AutoExtend := TRUE, Permissive := FALSE, FbRetracted := TRUE);
ASSERT_FALSE(c.Extend);
ASSERT_TRUE(c.Retract);
c(Mode := RB_MODE#Auto, AutoExtend := TRUE, Permissive := TRUE, FbRetracted := TRUE);
ASSERT_TRUE(c.Extend);
c(Mode := RB_MODE#Auto, AutoExtend := TRUE, Permissive := FALSE, FbExtended := TRUE, FbRetracted := FALSE);
ASSERT_TRUE(c.Extend);
END_TEST

TEST cylinder_stroke_faults
VAR a : RB_Cylinder; b : RB_Cylinder; k : RB_Cylinder; END_VAR
(* does not extend *)
a(Mode := RB_MODE#Auto, AutoExtend := TRUE, FbExtended := FALSE, FbRetracted := TRUE, MoveTime := T#1s);
ADVANCE(T#900ms);
a(Mode := RB_MODE#Auto, AutoExtend := TRUE, FbExtended := FALSE, FbRetracted := TRUE, MoveTime := T#1s);
ASSERT_FALSE(a.Error);
ADVANCE(T#200ms);
a(Mode := RB_MODE#Auto, AutoExtend := TRUE, FbExtended := FALSE, FbRetracted := TRUE, MoveTime := T#1s);
ASSERT_TRUE(a.Error);
ASSERT_EQ(UDINT#1, a.ErrorID);
ASSERT_FALSE(a.Extend);
ASSERT_FALSE(a.Retract);
ASSERT_EQ(UDINT#1, a.Status.ErrorID);
a(Mode := RB_MODE#Auto, AutoExtend := FALSE, FbExtended := FALSE, FbRetracted := TRUE, MoveTime := T#1s, Reset := TRUE);
ASSERT_FALSE(a.Error);
ASSERT_EQ(UDINT#0, a.ErrorID);
ASSERT_TRUE(a.Retract);
(* does not retract *)
b(Mode := RB_MODE#Auto, AutoExtend := FALSE, FbExtended := TRUE, FbRetracted := FALSE, MoveTime := T#1s);
ADVANCE(T#1100ms);
b(Mode := RB_MODE#Auto, AutoExtend := FALSE, FbExtended := TRUE, FbRetracted := FALSE, MoveTime := T#1s);
ASSERT_TRUE(b.Error);
ASSERT_EQ(UDINT#2, b.ErrorID);
(* both end switches *)
k(Mode := RB_MODE#Auto, AutoExtend := TRUE, FbExtended := TRUE, FbRetracted := TRUE, MoveTime := T#1s);
ASSERT_FALSE(k.IsExtended);
ASSERT_FALSE(k.IsRetracted);
ADVANCE(T#1100ms);
k(Mode := RB_MODE#Auto, AutoExtend := TRUE, FbExtended := TRUE, FbRetracted := TRUE, MoveTime := T#1s);
ASSERT_TRUE(k.Error);
ASSERT_EQ(UDINT#3, k.ErrorID);
END_TEST

TEST cylinder_single_acting_spring_return
VAR c : RB_Cylinder; d : RB_Cylinder; END_VAR
c(Mode := RB_MODE#Auto, AutoExtend := FALSE, DoubleActing := FALSE, FbExtended := FALSE, FbRetracted := TRUE, MoveTime := T#1s);
ASSERT_FALSE(c.Retract);
ASSERT_FALSE(c.Extend);
c(Mode := RB_MODE#Auto, AutoExtend := TRUE, DoubleActing := FALSE, FbExtended := FALSE, FbRetracted := TRUE, MoveTime := T#1s);
ASSERT_TRUE(c.Extend);
ASSERT_FALSE(c.Retract);
(* the spring does not bring it back in time *)
d(Mode := RB_MODE#Auto, AutoExtend := FALSE, DoubleActing := FALSE, FbExtended := TRUE, FbRetracted := FALSE, MoveTime := T#1s);
ADVANCE(T#1100ms);
d(Mode := RB_MODE#Auto, AutoExtend := FALSE, DoubleActing := FALSE, FbExtended := TRUE, FbRetracted := FALSE, MoveTime := T#1s);
ASSERT_TRUE(d.Error);
ASSERT_EQ(UDINT#2, d.ErrorID);
(* in Off the spring-return cylinder is not supervised for retracting *)
c(Mode := RB_MODE#Off, AutoExtend := FALSE, DoubleActing := FALSE, FbExtended := TRUE, FbRetracted := FALSE, MoveTime := T#1s);
ADVANCE(T#2s);
c(Mode := RB_MODE#Off, AutoExtend := FALSE, DoubleActing := FALSE, FbExtended := TRUE, FbRetracted := FALSE, MoveTime := T#1s);
ASSERT_FALSE(c.Error);
END_TEST

TEST cylinder_without_feedback
VAR c : RB_Cylinder; END_VAR
c(Mode := RB_MODE#Auto, AutoExtend := TRUE, Feedback := FALSE, FbExtended := FALSE, FbRetracted := TRUE, MoveTime := T#1s);
ASSERT_TRUE(c.IsExtended);
ASSERT_FALSE(c.IsRetracted);
ADVANCE(T#5s);
c(Mode := RB_MODE#Auto, AutoExtend := TRUE, Feedback := FALSE, FbExtended := TRUE, FbRetracted := TRUE, MoveTime := T#1s);
ASSERT_FALSE(c.Error);
c(Mode := RB_MODE#Auto, AutoExtend := TRUE, Feedback := TRUE, FbExtended := TRUE, FbRetracted := TRUE, MoveTime := T#1s);
ASSERT_FALSE(c.Error);
c(Mode := RB_MODE#Auto, AutoExtend := FALSE, Feedback := FALSE, FbExtended := FALSE, FbRetracted := TRUE, MoveTime := T#1s);
ASSERT_TRUE(c.IsRetracted);
END_TEST

TEST cylinder_supervision_switched_on_mid_stroke_starts_fresh
VAR c : RB_Cylinder; END_VAR
c(Mode := RB_MODE#Auto, AutoExtend := TRUE, Feedback := FALSE, FbExtended := FALSE, FbRetracted := FALSE, MoveTime := T#1s);
ADVANCE(T#5s);
c(Mode := RB_MODE#Auto, AutoExtend := TRUE, Feedback := FALSE, FbExtended := FALSE, FbRetracted := FALSE, MoveTime := T#1s);
c(Mode := RB_MODE#Auto, AutoExtend := TRUE, Feedback := TRUE, FbExtended := FALSE, FbRetracted := FALSE, MoveTime := T#1s);
ASSERT_FALSE(c.Error);
ADVANCE(T#1100ms);
c(Mode := RB_MODE#Auto, AutoExtend := TRUE, Feedback := TRUE, FbExtended := FALSE, FbRetracted := FALSE, MoveTime := T#1s);
ASSERT_TRUE(c.Error);
ASSERT_EQ(UDINT#1, c.ErrorID);
END_TEST

(* ---- ok_rb_data_logic.st ---- *)
(* spec: [blocks.fault] [blocks.interlock] [blocks.testable]
   expect: ok
   libraries: RootBlocks *)
(* Test suites of RB_Fifo (F11.FIFO), RB_RecipeTable (F11.RECIPE),
   RB_Transfer (F11.TRANSFER), RB_StartStop (F02.STARTSTOP) and
   RB_Permissives (F02.PERMISSIVES). Every call passes the inputs that
   matter: block inputs keep their last value. *)
TEST fifo_first_in_first_out
VAR q : RB_Fifo; END_VAR
q();
ASSERT_TRUE(q.Empty);
ASSERT_EQ(DINT#0, q.First);
q(Put := TRUE, InValue := 11);
q(Put := FALSE);
q(Put := TRUE, InValue := 22);
q(Put := FALSE);
ASSERT_EQ(2, q.Count);
ASSERT_EQ(DINT#11, q.First);
ASSERT_FALSE(q.Empty);
q(Get := TRUE);
ASSERT_EQ(DINT#11, q.OutValue);
ASSERT_EQ(DINT#22, q.First);
q(Get := FALSE);
q(Get := TRUE);
ASSERT_EQ(DINT#22, q.OutValue);
ASSERT_TRUE(q.Empty);
ASSERT_FALSE(q.Error);
(* a put and a get in the same call: the get takes the old value first *)
q(Get := FALSE, Put := TRUE, InValue := 33);
q(Put := FALSE);
q(Put := TRUE, Get := TRUE, InValue := 44);
ASSERT_EQ(DINT#33, q.OutValue);
ASSERT_EQ(1, q.Count);
ASSERT_EQ(DINT#44, q.First);
END_TEST

TEST fifo_wraps_and_reports_full_and_empty
VAR q : RB_Fifo; i : INT; END_VAR
FOR i := 1 TO 32 DO
    q(Put := TRUE, InValue := INT_TO_DINT(i));
    q(Put := FALSE);
END_FOR;
ASSERT_TRUE(q.Full);
q(Put := TRUE, InValue := 99);
ASSERT_TRUE(q.Error);
ASSERT_EQ(UDINT#1, q.ErrorID);
ASSERT_EQ(32, q.Count);
q(Put := FALSE, Reset := TRUE);
ASSERT_FALSE(q.Error);
ASSERT_EQ(UDINT#0, q.ErrorID);
(* take 5, put 5 more: the ring wraps around *)
FOR i := 1 TO 5 DO
    q(Get := TRUE, Reset := FALSE);
    q(Get := FALSE);
END_FOR;
ASSERT_EQ(DINT#5, q.OutValue);
FOR i := 1 TO 5 DO
    q(Put := TRUE, InValue := INT_TO_DINT(100 + i));
    q(Put := FALSE);
END_FOR;
FOR i := 1 TO 27 DO
    q(Get := TRUE);
    q(Get := FALSE);
END_FOR;
ASSERT_EQ(DINT#32, q.OutValue);
ASSERT_EQ(DINT#101, q.First);
q(Clear := TRUE);
ASSERT_TRUE(q.Empty);
ASSERT_FALSE(q.Full);
q(Clear := FALSE, Get := TRUE);
ASSERT_TRUE(q.Error);
ASSERT_EQ(UDINT#2, q.ErrorID);
END_TEST

TEST recipe_save_and_load
VAR r : RB_RecipeTable; t : ARRAY[1..16, 1..8] OF REAL; a : ARRAY[1..8] OF REAL; END_VAR
a[1] := 1.5;
a[8] := 8.5;
r(Number := 3, Save := TRUE, Actual := a, Table := t);
ASSERT_TRUE(r.Done);
ASSERT_TRUE(ABS(t[3, 1] - 1.5) < 0.0001);
ASSERT_TRUE(ABS(t[3, 8] - 8.5) < 0.0001);
ASSERT_EQ(0, r.Loaded);
r(Number := 3, Save := FALSE, Actual := a, Table := t);
ASSERT_FALSE(r.Done);
t[5, 2] := 42.0;
r(Number := 5, Load := TRUE, Table := t);
ASSERT_TRUE(r.Done);
ASSERT_EQ(5, r.Loaded);
ASSERT_TRUE(ABS(r.Params[2] - 42.0) < 0.0001);
ASSERT_TRUE(ABS(r.Params[1]) < 0.0001);
(* a save does not change the loaded parameters *)
r(Number := 3, Load := FALSE, Table := t);
r(Number := 3, Save := TRUE, Actual := a, Table := t);
ASSERT_TRUE(ABS(r.Params[2] - 42.0) < 0.0001);
ASSERT_EQ(5, r.Loaded);
END_TEST

TEST recipe_number_out_of_range
VAR r : RB_RecipeTable; t : ARRAY[1..16, 1..8] OF REAL; END_VAR
r(Number := 0, Load := TRUE, Table := t);
ASSERT_TRUE(r.Error);
ASSERT_EQ(UDINT#1, r.ErrorID);
ASSERT_FALSE(r.Done);
r(Number := 17, Load := FALSE, Reset := TRUE, Table := t);
ASSERT_FALSE(r.Error);
ASSERT_EQ(UDINT#0, r.ErrorID);
r(Number := 17, Save := TRUE, Reset := FALSE, Table := t);
ASSERT_TRUE(r.Error);
r(Number := 16, Save := FALSE, Reset := TRUE, Table := t);
r(Number := 16, Load := TRUE, Reset := FALSE, Table := t);
ASSERT_FALSE(r.Error);
ASSERT_EQ(16, r.Loaded);
r(Number := 1, Load := FALSE, Table := t);
r(Number := 1, Load := TRUE, Table := t);
ASSERT_EQ(1, r.Loaded);
END_TEST

TEST transfer_hands_a_part_on
VAR x : RB_Transfer; END_VAR
x(PartReady := TRUE, ReceiverReady := FALSE);
ASSERT_FALSE(x.Release);
x(PartReady := TRUE, ReceiverReady := TRUE);
ASSERT_TRUE(x.Release);
ASSERT_TRUE(x.Busy);
(* the receiver is busy now; the transfer goes on until arrival *)
x(PartReady := TRUE, ReceiverReady := FALSE, Arrived := FALSE);
ASSERT_TRUE(x.Release);
x(PartReady := FALSE, ReceiverReady := FALSE, Arrived := TRUE);
ASSERT_FALSE(x.Release);
ASSERT_TRUE(x.Done);
ASSERT_EQ(UDINT#1, x.Count);
x(PartReady := FALSE, ReceiverReady := TRUE, Arrived := TRUE);
ASSERT_FALSE(x.Done);
ASSERT_FALSE(x.Release);
ASSERT_FALSE(x.Busy);
END_TEST

TEST transfer_timeout
VAR x : RB_Transfer; END_VAR
x(PartReady := TRUE, ReceiverReady := TRUE, Timeout := T#2s);
ADVANCE(T#1900ms);
x(PartReady := TRUE, ReceiverReady := TRUE, Timeout := T#2s);
ASSERT_TRUE(x.Release);
ADVANCE(T#200ms);
x(PartReady := TRUE, ReceiverReady := TRUE, Timeout := T#2s);
ASSERT_TRUE(x.Error);
ASSERT_EQ(UDINT#1, x.ErrorID);
ASSERT_FALSE(x.Release);
(* no new transfer while the error lasts *)
x(PartReady := TRUE, ReceiverReady := TRUE, Timeout := T#2s);
ASSERT_FALSE(x.Release);
x(PartReady := TRUE, ReceiverReady := TRUE, Timeout := T#2s, Reset := TRUE);
ASSERT_FALSE(x.Error);
ASSERT_EQ(UDINT#0, x.ErrorID);
ASSERT_TRUE(x.Release);
END_TEST

TEST start_stop_latch_stop_wins
VAR s : RB_StartStop; END_VAR
s(Start := TRUE);
ASSERT_TRUE(s.Out);
s(Start := FALSE);
ASSERT_TRUE(s.Out);
s(StopOk := FALSE);
ASSERT_FALSE(s.Out);
(* start while stop is pressed: stop wins *)
s(Start := TRUE, StopOk := FALSE);
ASSERT_FALSE(s.Out);
s(Start := FALSE, StopOk := TRUE);
ASSERT_FALSE(s.Out);
s(Start := TRUE, Permissive := FALSE);
ASSERT_FALSE(s.Out);
s(Start := FALSE, Permissive := TRUE);
s(Start := TRUE);
ASSERT_TRUE(s.Out);
s(Permissive := FALSE);
ASSERT_TRUE(s.Out);
s(Interlock := TRUE);
ASSERT_FALSE(s.Out);
END_TEST

TEST permissives_and_first_out
VAR p : RB_Permissives; c : ARRAY[1..16] OF BOOL; k : INT; END_VAR
FOR k := 1 TO 16 DO c[k] := TRUE; END_FOR;
p(Cond := c);
ASSERT_TRUE(p.Ok);
ASSERT_EQ(0, p.FirstOut);
c[7] := FALSE;
p(Cond := c);
ASSERT_FALSE(p.Ok);
ASSERT_EQ(7, p.FirstOut);
ASSERT_EQ(1, p.Missing);
c[3] := FALSE;
p(Cond := c);
ASSERT_EQ(7, p.FirstOut);
ASSERT_EQ(2, p.Missing);
(* reset only clears when all are back *)
p(Cond := c, Reset := TRUE);
ASSERT_EQ(7, p.FirstOut);
c[3] := TRUE;
c[7] := TRUE;
p(Cond := c, Reset := FALSE);
ASSERT_TRUE(p.Ok);
ASSERT_EQ(7, p.FirstOut);
p(Cond := c, Reset := TRUE);
ASSERT_EQ(0, p.FirstOut);
(* unused conditions do not count *)
c[16] := FALSE;
c[1] := FALSE;
p(Cond := c, Reset := FALSE, Used := WORD#16#7FFE);
ASSERT_TRUE(p.Ok);
p(Cond := c, Used := WORD#16#FFFF);
ASSERT_EQ(1, p.FirstOut);
ASSERT_EQ(2, p.Missing);
END_TEST

(* ---- ok_rb_devices2.st ---- *)
(* spec: [blocks.mode] [blocks.interlock] [blocks.fault] [blocks.feedback] [blocks.status] [blocks.testable]
   expect: ok
   libraries: RootBlocks *)
(* Test suites of RB_ValveAnalog (F04.VALVE.ANALOG), RB_MotorStarDelta
   (F04.MOTOR.STARDELTA) and RB_Diverter (F12.DIVERTER). Every call passes
   the inputs that matter: block inputs keep their last value. *)
TEST valve_analog_modes_and_limits
VAR v : RB_ValveAnalog; END_VAR
v(Mode := RB_MODE#Off, AutoPos := 40.0, ManPos := 70.0, Feedback := FALSE);
ASSERT_TRUE(ABS(v.Out) < 0.001);
ASSERT_FALSE(v.Status.Commanded);
v(Mode := RB_MODE#Auto);
ASSERT_TRUE(ABS(v.Out - 40.0) < 0.001);
ASSERT_TRUE(ABS(v.Pos - 40.0) < 0.001);
ASSERT_TRUE(v.Status.Commanded);
ASSERT_TRUE(v.Status.Active);
ASSERT_EQ(UDINT#1, v.Status.Starts);
v(Mode := RB_MODE#Manual);
ASSERT_TRUE(ABS(v.Out - 70.0) < 0.001);
ASSERT_EQ(UDINT#1, v.Status.Starts);
ASSERT_TRUE(v.Status.Mode = RB_MODE#Manual);
v(ManPos := 120.0);
ASSERT_TRUE(ABS(v.Out - 100.0) < 0.001);
v(ManPos := -5.0);
ASSERT_TRUE(ABS(v.Out) < 0.001);
ASSERT_FALSE(v.Status.Active);
v(ManPos := 3.0);
ASSERT_EQ(UDINT#2, v.Status.Starts);
(* a small opening is not reported as open (below Tolerance) *)
ASSERT_FALSE(v.Status.Active);
v(ManPos := 5.0);
ASSERT_FALSE(v.Status.Active);
v(ManPos := 6.0);
ASSERT_TRUE(v.Status.Active);
END_TEST

TEST valve_analog_interlock_goes_to_the_safe_position
VAR v : RB_ValveAnalog; END_VAR
v(Mode := RB_MODE#Auto, AutoPos := 40.0, Feedback := FALSE);
v(Interlock := TRUE);
ASSERT_TRUE(ABS(v.Out) < 0.001);
(* a valve that must open on a fault *)
v(SafePos := 100.0);
ASSERT_TRUE(ABS(v.Out - 100.0) < 0.001);
v(Interlock := FALSE);
ASSERT_TRUE(ABS(v.Out - 40.0) < 0.001);
v(Mode := RB_MODE#Off);
ASSERT_TRUE(ABS(v.Out - 100.0) < 0.001);
END_TEST

TEST valve_analog_deviation_fault
VAR v : RB_ValveAnalog; END_VAR
v(Mode := RB_MODE#Auto, AutoPos := 50.0, PosFb := 0.0, FeedbackTime := T#2s);
ASSERT_TRUE(ABS(v.Pos) < 0.001);
ADVANCE(T#1900ms);
v(PosFb := 30.0);
ASSERT_FALSE(v.Error);
ASSERT_TRUE(ABS(v.Pos - 30.0) < 0.001);
(* within tolerance: the timer restarts *)
v(PosFb := 45.0);
ADVANCE(T#5s);
v(PosFb := 45.0);
ASSERT_FALSE(v.Error);
v(PosFb := 44.0);
ADVANCE(T#1900ms);
v(PosFb := 44.0);
ASSERT_FALSE(v.Error);
ADVANCE(T#200ms);
v(PosFb := 44.0);
ASSERT_TRUE(v.Error);
ASSERT_EQ(UDINT#1, v.ErrorID);
ASSERT_TRUE(ABS(v.Out) < 0.001);
ASSERT_TRUE(v.Status.Error);
ASSERT_EQ(UDINT#1, v.Status.ErrorID);
(* the fault holds the safe position until reset *)
v(PosFb := 0.0);
ASSERT_TRUE(ABS(v.Out) < 0.001);
v(PosFb := 0.0, Reset := TRUE);
ASSERT_FALSE(v.Error);
ASSERT_EQ(UDINT#0, v.ErrorID);
ASSERT_TRUE(ABS(v.Out - 50.0) < 0.001);
END_TEST

TEST valve_analog_feedback_out_of_range
VAR v : RB_ValveAnalog; END_VAR
v(Mode := RB_MODE#Auto, AutoPos := 50.0, PosFb := 110.0);
ASSERT_FALSE(v.Error);
v(PosFb := 111.0);
ASSERT_TRUE(v.Error);
ASSERT_EQ(UDINT#2, v.ErrorID);
v(PosFb := 50.0, Reset := TRUE);
ASSERT_FALSE(v.Error);
v(PosFb := -10.0, Reset := FALSE);
ASSERT_FALSE(v.Error);
v(PosFb := -11.0);
ASSERT_TRUE(v.Error);
ASSERT_EQ(UDINT#2, v.ErrorID);
(* without feedback the signal is ignored *)
v(PosFb := -50.0, Reset := TRUE, Feedback := FALSE);
ASSERT_FALSE(v.Error);
ADVANCE(T#20s);
v(PosFb := -50.0, Reset := FALSE);
ASSERT_FALSE(v.Error);
ASSERT_TRUE(ABS(v.Pos - 50.0) < 0.001);
(* switching supervision back on starts the timer fresh *)
v(PosFb := 0.0, Feedback := TRUE);
ADVANCE(T#9s);
v(PosFb := 0.0, Feedback := FALSE);
v(PosFb := 0.0, Feedback := TRUE);
ADVANCE(T#2s);
v(PosFb := 0.0);
ASSERT_FALSE(v.Error);
END_TEST

TEST star_delta_starts_in_star_then_delta
VAR m : RB_MotorStarDelta; END_VAR
m(Mode := RB_MODE#Auto, AutoRun := FALSE);
ASSERT_FALSE(m.Main OR m.Star OR m.Delta);
m(AutoRun := TRUE, FbRunning := FALSE);
ASSERT_TRUE(m.Main);
ASSERT_TRUE(m.Star);
ASSERT_FALSE(m.Delta);
ASSERT_FALSE(m.Running);
ASSERT_EQ(UDINT#1, m.Status.Starts);
ADVANCE(T#4900ms);
m(FbRunning := TRUE);
ASSERT_TRUE(m.Star);
ASSERT_TRUE(m.Running);
ASSERT_FALSE(m.InDelta);
(* star off, a short gap with both off, then delta *)
ADVANCE(T#100ms);
m();
ASSERT_TRUE(m.Main);
ASSERT_FALSE(m.Star);
ASSERT_FALSE(m.Delta);
ADVANCE(T#40ms);
m();
ASSERT_FALSE(m.Delta);
ADVANCE(T#10ms);
m();
ASSERT_TRUE(m.Delta);
ASSERT_TRUE(m.InDelta);
ASSERT_FALSE(m.Star);
ADVANCE(T#10s);
m();
ASSERT_TRUE(m.Delta);
(* stop and start again: star first *)
m(AutoRun := FALSE, FbRunning := TRUE);
ASSERT_FALSE(m.Main OR m.Star OR m.Delta);
m(AutoRun := TRUE);
ASSERT_TRUE(m.Star);
ASSERT_FALSE(m.Delta);
ASSERT_EQ(UDINT#2, m.Status.Starts);
END_TEST

TEST star_delta_faults_and_settings
VAR m : RB_MotorStarDelta; END_VAR
m(Mode := RB_MODE#Manual, ManRun := TRUE, FbRunning := TRUE, StarTime := T#2s, Changeover := T#100ms);
ASSERT_TRUE(m.Star);
ADVANCE(T#2s);
m();
ASSERT_FALSE(m.Star);
ADVANCE(T#100ms);
m();
ASSERT_TRUE(m.Delta);
m(Overload := TRUE);
ASSERT_TRUE(m.Error);
ASSERT_EQ(UDINT#3, m.ErrorID);
ASSERT_FALSE(m.Main OR m.Star OR m.Delta);
ASSERT_TRUE(m.Status.Error);
m(Overload := FALSE, Reset := TRUE, FbRunning := FALSE);
ASSERT_FALSE(m.Error);
ASSERT_TRUE(m.Star);
(* no running feedback: fault 1 *)
ADVANCE(T#3s);
m(Reset := FALSE, FeedbackTime := T#2s);
ASSERT_TRUE(m.Error);
ASSERT_EQ(UDINT#1, m.ErrorID);
(* interlock, permissive, restart delay pass through RB_Motor *)
m(Reset := TRUE, Feedback := FALSE, Interlock := TRUE);
ASSERT_FALSE(m.Main);
m(Reset := FALSE, Interlock := FALSE, ManRun := FALSE);
m(ManRun := TRUE, Permissive := FALSE);
ASSERT_FALSE(m.Main);
m(ManRun := TRUE, Permissive := TRUE, RestartDelay := T#1s);
ASSERT_FALSE(m.Main);
ADVANCE(T#1s);
m();
ASSERT_TRUE(m.Main);
ASSERT_TRUE(m.Running);
END_TEST

TEST diverter_sends_a_part_into_the_branch
VAR d : RB_Diverter; END_VAR
d(FbStraight := TRUE);
ASSERT_FALSE(d.Gate);
ASSERT_FALSE(d.HoldPart);
(* the part arrives for the branch: hold it until the gate is over *)
d(PartAtGate := TRUE, Divert := TRUE, FbStraight := TRUE);
ASSERT_TRUE(d.Gate);
ASSERT_TRUE(d.HoldPart);
d(PartAtGate := TRUE, Divert := FALSE, FbStraight := FALSE, FbDiverted := TRUE);
ASSERT_TRUE(d.Gate);
ASSERT_FALSE(d.HoldPart);
(* it leaves the eye: counted, the gate stays for PassTime *)
d(PartAtGate := FALSE);
ASSERT_EQ(UDINT#1, d.ToBranch);
ASSERT_EQ(UDINT#0, d.ToStraight);
ADVANCE(T#900ms);
d();
ASSERT_TRUE(d.Gate);
ADVANCE(T#100ms);
d();
ASSERT_FALSE(d.Gate);
(* the gate swings back; no part is waiting, nothing to hold *)
ASSERT_FALSE(d.HoldPart);
d(FbDiverted := FALSE, FbStraight := TRUE);
ASSERT_FALSE(d.Error);
END_TEST

TEST diverter_straight_parts_and_a_quick_follower
VAR d : RB_Diverter; END_VAR
d(PartAtGate := TRUE, Divert := FALSE, FbStraight := TRUE);
ASSERT_FALSE(d.Gate);
ASSERT_FALSE(d.HoldPart);
d(PartAtGate := FALSE);
ASSERT_EQ(UDINT#1, d.ToStraight);
(* the next part, for the branch, comes during PassTime *)
ADVANCE(T#300ms);
d(PartAtGate := TRUE, Divert := TRUE);
ASSERT_TRUE(d.Gate);
ASSERT_TRUE(d.HoldPart);
ADVANCE(T#900ms);
d(FbStraight := FALSE, FbDiverted := TRUE);
ASSERT_TRUE(d.Gate);
ASSERT_FALSE(d.HoldPart);
d(PartAtGate := FALSE);
ASSERT_EQ(UDINT#1, d.ToBranch);
(* both gate switches on: not in position, the part is held *)
d(PartAtGate := FALSE);
ADVANCE(T#2s);
d(PartAtGate := FALSE, FbStraight := TRUE, FbDiverted := TRUE);
d(PartAtGate := TRUE, Divert := FALSE);
ASSERT_TRUE(d.HoldPart);
d(PartAtGate := FALSE, FbDiverted := FALSE);
ASSERT_EQ(UDINT#2, d.ToStraight);
ADVANCE(T#2s);
d();
(* a part leaving without arriving (power-up) is not counted *)
d(PartAtGate := TRUE, Divert := FALSE);
ADVANCE(T#5s);
d(PartAtGate := TRUE, FbStraight := TRUE, FbDiverted := FALSE);
d(PartAtGate := FALSE);
ASSERT_EQ(UDINT#3, d.ToStraight);
END_TEST

TEST diverter_gate_timeout
VAR d : RB_Diverter; END_VAR
d(PartAtGate := TRUE, Divert := TRUE, FbStraight := TRUE, MoveTime := T#1s);
ADVANCE(T#900ms);
d();
ASSERT_FALSE(d.Error);
ADVANCE(T#100ms);
d();
ASSERT_TRUE(d.Error);
ASSERT_EQ(UDINT#1, d.ErrorID);
ASSERT_FALSE(d.Gate);
ASSERT_TRUE(d.HoldPart);
(* the gate is straight again: reset; the part still waits, the gate retries *)
d(Reset := TRUE);
ASSERT_FALSE(d.Error);
ASSERT_EQ(UDINT#0, d.ErrorID);
ASSERT_TRUE(d.Gate);
d(Reset := FALSE, FbStraight := FALSE, FbDiverted := TRUE);
ASSERT_FALSE(d.HoldPart);
(* both switches on: not in position *)
d(FbStraight := TRUE, FbDiverted := TRUE);
ASSERT_TRUE(d.HoldPart);
END_TEST

TEST diverter_without_feedback
VAR d : RB_Diverter; END_VAR
d(Feedback := FALSE, PartAtGate := TRUE, Divert := TRUE);
ASSERT_TRUE(d.Gate);
ASSERT_FALSE(d.HoldPart);
ADVANCE(T#10s);
d();
ASSERT_FALSE(d.Error);
END_TEST

(* ---- ok_rb_drive.st ---- *)
(* spec: [blocks.command] [blocks.mode] [blocks.interlock] [blocks.fault] [blocks.feedback] [blocks.status]
   expect: ok
   libraries: RootBlocks *)
(* Test suite of RB_Drive (card blocks/cards/F04.DRIVE.md). Every call passes
   the inputs that matter: block inputs keep their last value. *)
TEST drive_runs_at_the_clamped_set_point
VAR d : RB_Drive; END_VAR
d(Mode := RB_MODE#Auto, AutoRun := TRUE, AutoSpeed := 60.0, DriveReady := TRUE, DriveRunning := FALSE);
ASSERT_TRUE(d.Run);
ASSERT_TRUE(ABS(d.SpeedSetpoint - 60.0) < 0.001);
ASSERT_FALSE(d.Reverse);
ASSERT_FALSE(d.Running);
ASSERT_FALSE(d.AtSpeed);
d(Mode := RB_MODE#Auto, AutoRun := TRUE, AutoSpeed := 130.0, DriveReady := TRUE, DriveRunning := TRUE);
ASSERT_TRUE(ABS(d.SpeedSetpoint - 100.0) < 0.001);
ASSERT_TRUE(d.Running);
ASSERT_TRUE(d.AtSpeed);
ASSERT_TRUE(d.Status.Active);
ASSERT_TRUE(d.Status.Commanded);
ASSERT_EQ(UDINT#1, d.Status.Starts);
ASSERT_TRUE(d.Status.Mode = RB_MODE#Auto);
d(Mode := RB_MODE#Auto, AutoRun := TRUE, AutoSpeed := 5.0, SpeedMin := 20.0, AutoReverse := TRUE, DriveReady := TRUE, DriveRunning := TRUE);
ASSERT_TRUE(ABS(d.SpeedSetpoint - 20.0) < 0.001);
ASSERT_TRUE(d.Reverse);
ASSERT_EQ(UDINT#1, d.Status.Starts);
d(Mode := RB_MODE#Auto, AutoRun := FALSE, AutoSpeed := 50.0, AutoReverse := TRUE, DriveReady := TRUE, DriveRunning := TRUE);
ASSERT_FALSE(d.Run);
ASSERT_TRUE(ABS(d.SpeedSetpoint) < 0.001);
ASSERT_FALSE(d.Reverse);
ASSERT_FALSE(d.Error);
ASSERT_FALSE(d.Status.Error);
END_TEST

TEST drive_modes_interlock_permissive_ready
VAR d : RB_Drive; END_VAR
d(Mode := RB_MODE#Auto, ManRun := TRUE, ManSpeed := 30.0, DriveReady := TRUE);
ASSERT_FALSE(d.Run);
d(Mode := RB_MODE#Manual, ManRun := TRUE, ManSpeed := 30.0, ManReverse := TRUE, AutoRun := FALSE, DriveReady := TRUE);
ASSERT_TRUE(d.Run);
ASSERT_TRUE(ABS(d.SpeedSetpoint - 30.0) < 0.001);
ASSERT_TRUE(d.Reverse);
d(Mode := RB_MODE#Manual, ManRun := TRUE, Interlock := TRUE, DriveReady := TRUE, DriveRunning := TRUE);
ASSERT_FALSE(d.Run);
d(Mode := RB_MODE#Off, ManRun := TRUE, AutoRun := TRUE, AutoSpeed := 40.0, AutoReverse := TRUE, Interlock := FALSE, DriveReady := TRUE, DriveRunning := FALSE);
ASSERT_FALSE(d.Run);
ASSERT_FALSE(d.Reverse);
ASSERT_TRUE(ABS(d.SpeedSetpoint) < 0.001);
d(Mode := RB_MODE#Auto, AutoRun := TRUE, Permissive := FALSE, DriveReady := TRUE, DriveRunning := FALSE);
ASSERT_FALSE(d.Run);
d(Mode := RB_MODE#Auto, AutoRun := TRUE, Permissive := TRUE, DriveReady := FALSE, DriveRunning := FALSE);
ASSERT_FALSE(d.Run);
d(Mode := RB_MODE#Auto, AutoRun := TRUE, Permissive := TRUE, DriveReady := TRUE, DriveRunning := FALSE);
ASSERT_TRUE(d.Run);
d(Mode := RB_MODE#Auto, AutoRun := TRUE, Permissive := FALSE, DriveReady := FALSE, DriveRunning := TRUE);
ASSERT_TRUE(d.Run);
END_TEST

TEST drive_fault_from_the_drive_and_reset_pulse
VAR d : RB_Drive; END_VAR
d(Mode := RB_MODE#Auto, AutoRun := TRUE, AutoSpeed := 50.0, AutoReverse := TRUE, DriveReady := TRUE, DriveRunning := TRUE);
ASSERT_TRUE(d.Reverse);
d(Mode := RB_MODE#Auto, AutoRun := TRUE, AutoSpeed := 50.0, AutoReverse := TRUE, DriveReady := FALSE, DriveRunning := FALSE, DriveFault := TRUE);
ASSERT_FALSE(d.Reverse);
ASSERT_TRUE(d.Error);
ASSERT_EQ(UDINT#3, d.ErrorID);
ASSERT_FALSE(d.Run);
ASSERT_TRUE(ABS(d.SpeedSetpoint) < 0.001);
ASSERT_FALSE(d.ResetDrive);
d(Mode := RB_MODE#Auto, AutoRun := TRUE, DriveReady := TRUE, DriveFault := FALSE, Reset := TRUE);
ASSERT_TRUE(d.ResetDrive);
ASSERT_FALSE(d.Error);
ASSERT_EQ(UDINT#0, d.ErrorID);
ASSERT_TRUE(d.Run);
d(Mode := RB_MODE#Auto, AutoRun := TRUE, DriveReady := TRUE, DriveRunning := TRUE, Reset := TRUE);
ASSERT_FALSE(d.ResetDrive);
END_TEST

TEST drive_run_feedback_supervision
VAR a : RB_Drive; b : RB_Drive; END_VAR
a(Mode := RB_MODE#Auto, AutoRun := TRUE, AutoSpeed := 50.0, DriveReady := TRUE, DriveRunning := FALSE, FeedbackTime := T#1s);
ADVANCE(T#900ms);
a(Mode := RB_MODE#Auto, AutoRun := TRUE, AutoSpeed := 50.0, DriveReady := TRUE, DriveRunning := FALSE, FeedbackTime := T#1s);
ASSERT_FALSE(a.Error);
ADVANCE(T#200ms);
a(Mode := RB_MODE#Auto, AutoRun := TRUE, AutoSpeed := 50.0, DriveReady := TRUE, DriveRunning := FALSE, FeedbackTime := T#1s);
ASSERT_TRUE(a.Error);
ASSERT_EQ(UDINT#1, a.ErrorID);
ASSERT_EQ(UDINT#1, a.Status.ErrorID);
b(Mode := RB_MODE#Auto, AutoRun := FALSE, DriveReady := TRUE, DriveRunning := TRUE, FeedbackTime := T#1s);
ADVANCE(T#1100ms);
b(Mode := RB_MODE#Auto, AutoRun := FALSE, DriveReady := TRUE, DriveRunning := TRUE, FeedbackTime := T#1s);
ASSERT_TRUE(b.Error);
ASSERT_EQ(UDINT#2, b.ErrorID);
END_TEST

TEST drive_speed_deviation
VAR d : RB_Drive; e : RB_Drive; END_VAR
d(Mode := RB_MODE#Auto, AutoRun := TRUE, AutoSpeed := 50.0, DriveReady := TRUE, DriveRunning := TRUE, ActualSpeed := 50.0, SpeedTolerance := 2.0, FeedbackTime := T#1s);
ASSERT_TRUE(d.AtSpeed);
d(Mode := RB_MODE#Auto, AutoRun := TRUE, AutoSpeed := 50.0, DriveReady := TRUE, DriveRunning := TRUE, ActualSpeed := 52.0, SpeedTolerance := 2.0, FeedbackTime := T#1s);
ASSERT_TRUE(d.AtSpeed);
d(Mode := RB_MODE#Auto, AutoRun := TRUE, AutoSpeed := 50.0, DriveReady := TRUE, DriveRunning := TRUE, ActualSpeed := 40.0, SpeedTolerance := 2.0, FeedbackTime := T#1s);
ASSERT_FALSE(d.AtSpeed);
ADVANCE(T#900ms);
d(Mode := RB_MODE#Auto, AutoRun := TRUE, AutoSpeed := 50.0, DriveReady := TRUE, DriveRunning := TRUE, ActualSpeed := 40.0, SpeedTolerance := 2.0, FeedbackTime := T#1s);
ASSERT_FALSE(d.Error);
ADVANCE(T#200ms);
d(Mode := RB_MODE#Auto, AutoRun := TRUE, AutoSpeed := 50.0, DriveReady := TRUE, DriveRunning := TRUE, ActualSpeed := 40.0, SpeedTolerance := 2.0, FeedbackTime := T#1s);
ASSERT_TRUE(d.Error);
ASSERT_EQ(UDINT#4, d.ErrorID);
(* without a tolerance the speed is not supervised *)
e(Mode := RB_MODE#Auto, AutoRun := TRUE, AutoSpeed := 50.0, DriveReady := TRUE, DriveRunning := TRUE, ActualSpeed := 10.0, SpeedTolerance := 0.0, FeedbackTime := T#1s);
ADVANCE(T#3s);
e(Mode := RB_MODE#Auto, AutoRun := TRUE, AutoSpeed := 50.0, DriveReady := TRUE, DriveRunning := TRUE, ActualSpeed := 10.0, SpeedTolerance := 0.0, FeedbackTime := T#1s);
ASSERT_FALSE(e.Error);
ASSERT_TRUE(e.AtSpeed);
(* a running drive that is not commanded is no speed deviation *)
e(Mode := RB_MODE#Auto, AutoRun := FALSE, DriveReady := TRUE, DriveRunning := FALSE, ActualSpeed := 30.0, SpeedTolerance := 2.0, FeedbackTime := T#1s);
ADVANCE(T#3s);
e(Mode := RB_MODE#Auto, AutoRun := FALSE, DriveReady := TRUE, DriveRunning := FALSE, ActualSpeed := 30.0, SpeedTolerance := 2.0, FeedbackTime := T#1s);
ASSERT_FALSE(e.Error);
END_TEST

(* ---- ok_rb_handling.st ---- *)
(* spec: [blocks.fault] [blocks.testable]
   expect: ok
   libraries: RootBlocks *)
(* Test suites of RB_ConveyorZone (F12.ZONE), RB_RunHours (F09.RUNHOURS)
   and RB_Heartbeat (F09.HEARTBEAT). Every call passes the inputs that
   matter: block inputs keep their last value. *)
TEST zone_accumulates_and_hands_on
VAR z : RB_ConveyorZone; END_VAR
(* empty zone: runs to bring parts forward *)
z(Enable := TRUE, PartAtEnd := FALSE, DownstreamFree := FALSE);
ASSERT_TRUE(z.Run);
ASSERT_TRUE(z.Free);
ASSERT_FALSE(z.Occupied);
ASSERT_FALSE(z.Feeding);
(* a part arrives, the next zone is full: stop and wait *)
z(Enable := TRUE, PartAtEnd := TRUE, DownstreamFree := FALSE);
ASSERT_FALSE(z.Run);
ASSERT_TRUE(z.Occupied);
ASSERT_FALSE(z.Free);
(* the next zone is free: hand it on *)
z(Enable := TRUE, PartAtEnd := TRUE, DownstreamFree := TRUE);
ASSERT_TRUE(z.Run);
ASSERT_TRUE(z.Feeding);
z(Enable := TRUE, PartAtEnd := FALSE, DownstreamFree := TRUE);
ASSERT_EQ(UDINT#1, z.Count);
ASSERT_FALSE(z.Feeding);
ASSERT_TRUE(z.Run);
(* the line stops *)
z(Enable := FALSE, PartAtEnd := FALSE, DownstreamFree := TRUE);
ASSERT_FALSE(z.Run);
ASSERT_FALSE(z.Free);
z(Enable := FALSE, PartAtEnd := TRUE, DownstreamFree := TRUE);
ASSERT_FALSE(z.Feeding);
ASSERT_FALSE(z.Run);
(* a part removed by hand while stopped is not counted *)
z(Enable := FALSE, PartAtEnd := FALSE, DownstreamFree := TRUE);
ASSERT_EQ(UDINT#1, z.Count);
ASSERT_FALSE(z.Occupied);
END_TEST

TEST zone_is_occupied_from_the_hand_over
VAR z : RB_ConveyorZone; END_VAR
z(Enable := TRUE, PartAtEnd := FALSE, DownstreamFree := FALSE, UpstreamFeeding := FALSE);
ASSERT_TRUE(z.Free);
z(Enable := TRUE, PartAtEnd := FALSE, DownstreamFree := FALSE, UpstreamFeeding := TRUE);
ASSERT_TRUE(z.Free);
(* the previous zone has handed the part over: occupied, still travelling *)
z(Enable := TRUE, PartAtEnd := FALSE, DownstreamFree := FALSE, UpstreamFeeding := FALSE);
ASSERT_TRUE(z.Occupied);
ASSERT_FALSE(z.Free);
ASSERT_TRUE(z.Run);
z(Enable := TRUE, PartAtEnd := TRUE, DownstreamFree := FALSE, UpstreamFeeding := FALSE);
ASSERT_FALSE(z.Run);
ASSERT_TRUE(z.Occupied);
z(Enable := TRUE, PartAtEnd := TRUE, DownstreamFree := TRUE, UpstreamFeeding := FALSE);
z(Enable := TRUE, PartAtEnd := FALSE, DownstreamFree := TRUE, UpstreamFeeding := FALSE);
ASSERT_FALSE(z.Occupied);
ASSERT_TRUE(z.Free);
END_TEST

TEST zone_sleeps_when_empty_and_not_fed
VAR z : RB_ConveyorZone; END_VAR
z(Enable := TRUE, PartAtEnd := FALSE, SleepTime := T#10s);
ADVANCE(T#9s);
z(Enable := TRUE, PartAtEnd := FALSE, SleepTime := T#10s);
ASSERT_TRUE(z.Run);
ADVANCE(T#2s);
z(Enable := TRUE, PartAtEnd := FALSE, SleepTime := T#10s);
ASSERT_FALSE(z.Run);
ASSERT_TRUE(z.Free);
(* the previous zone feeds a part: wake up *)
z(Enable := TRUE, PartAtEnd := FALSE, UpstreamFeeding := TRUE, SleepTime := T#10s);
ASSERT_TRUE(z.Run);
(* without a sleep time it never stops *)
ADVANCE(T#1h);
z(Enable := TRUE, PartAtEnd := FALSE, UpstreamFeeding := FALSE, SleepTime := T#0s);
ASSERT_TRUE(z.Run);
END_TEST

TEST zone_jam_latches_until_reset
VAR z : RB_ConveyorZone; y : RB_ConveyorZone; END_VAR
z(Enable := TRUE, PartAtEnd := TRUE, DownstreamFree := TRUE, JamTime := T#2s);
ADVANCE(T#1900ms);
z(Enable := TRUE, PartAtEnd := TRUE, DownstreamFree := TRUE, JamTime := T#2s);
ASSERT_FALSE(z.Error);
ADVANCE(T#200ms);
z(Enable := TRUE, PartAtEnd := TRUE, DownstreamFree := TRUE, JamTime := T#2s);
ASSERT_TRUE(z.Error);
ASSERT_EQ(UDINT#1, z.ErrorID);
ASSERT_FALSE(z.Run);
ASSERT_FALSE(z.Feeding);
ASSERT_FALSE(z.Free);
(* the jam cleared by hand: still latched *)
z(Enable := TRUE, PartAtEnd := FALSE, DownstreamFree := TRUE, JamTime := T#2s);
ASSERT_TRUE(z.Error);
ASSERT_FALSE(z.Run);
z(Enable := TRUE, PartAtEnd := FALSE, DownstreamFree := TRUE, JamTime := T#2s, Reset := TRUE);
ASSERT_FALSE(z.Error);
ASSERT_EQ(UDINT#0, z.ErrorID);
ASSERT_TRUE(z.Run);
(* without jam supervision a part may wait as long as it likes *)
y(Enable := TRUE, PartAtEnd := TRUE, DownstreamFree := TRUE, JamTime := T#0s);
ADVANCE(T#1h);
y(Enable := TRUE, PartAtEnd := TRUE, DownstreamFree := TRUE, JamTime := T#0s);
ASSERT_FALSE(y.Error);
END_TEST

TEST run_hours_and_starts
VAR h : RB_RunHours; END_VAR
h(Running := FALSE, Interval := 2.0);
ADVANCE(T#1h);
h(Running := FALSE, Interval := 2.0);
ASSERT_TRUE(ABS(h.Hours) < 0.000001);
h(Running := TRUE, Interval := 2.0);
ASSERT_EQ(UDINT#1, h.Starts);
ADVANCE(T#90m);
h(Running := TRUE, Interval := 2.0);
ASSERT_TRUE(ABS(h.Hours - 1.5) < 0.0001);
ASSERT_FALSE(h.MaintenanceDue);
ADVANCE(T#30m);
h(Running := TRUE, Interval := 2.0);
ASSERT_TRUE(ABS(h.SinceService - 2.0) < 0.0001);
ASSERT_TRUE(h.MaintenanceDue);
h(Running := TRUE, Interval := 2.0);
ASSERT_EQ(UDINT#1, h.Starts);
h(Running := FALSE, Interval := 2.0, ServiceDone := TRUE);
ASSERT_TRUE(ABS(h.SinceService) < 0.0001);
ASSERT_FALSE(h.MaintenanceDue);
ASSERT_TRUE(ABS(h.Hours - 2.0) < 0.0001);
(* no interval: never due *)
h(Running := FALSE, Interval := 0.0);
ASSERT_FALSE(h.MaintenanceDue);
(* the time up to the call that sees the stop counts *)
h(Running := TRUE, Interval := 0.0);
ADVANCE(T#1h);
h(Running := FALSE, Interval := 0.0);
ASSERT_TRUE(ABS(h.Hours - 3.0) < 0.0001);
END_TEST

TEST run_hours_restored_from_a_preset
VAR h : RB_RunHours; END_VAR
h(Load := TRUE, PresetHours := 1000.0, PresetStarts := 42, PresetSince := 99.0, Interval := 100.0);
ASSERT_TRUE(ABS(h.Hours - 1000.0) < 0.0001);
ASSERT_EQ(UDINT#42, h.Starts);
ASSERT_FALSE(h.MaintenanceDue);
h(Load := TRUE, Running := TRUE, PresetHours := 0.0, Interval := 100.0);
ASSERT_TRUE(ABS(h.Hours - 1000.0) < 0.0001);
ASSERT_EQ(UDINT#43, h.Starts);
ADVANCE(T#1h);
h(Load := FALSE, Running := TRUE, Interval := 100.0);
ASSERT_TRUE(h.MaintenanceDue);
END_TEST

TEST heartbeat_toggles_and_supervises
VAR b : RB_Heartbeat; END_VAR
b(PartnerBeat := FALSE, Period := T#1s, Timeout := T#3s);
ASSERT_FALSE(b.Beat);
ASSERT_TRUE(b.Alive);
ADVANCE(T#1s);
b(PartnerBeat := TRUE, Period := T#1s, Timeout := T#3s);
ASSERT_TRUE(b.Beat);
ADVANCE(T#500ms);
b(PartnerBeat := TRUE, Period := T#1s, Timeout := T#3s);
ASSERT_TRUE(b.Beat);
ADVANCE(T#500ms);
b(PartnerBeat := FALSE, Period := T#1s, Timeout := T#3s);
ASSERT_FALSE(b.Beat);
ASSERT_TRUE(b.Alive);
(* the partner stops beating *)
ADVANCE(T#2900ms);
b(PartnerBeat := FALSE, Period := T#1s, Timeout := T#3s);
ASSERT_TRUE(b.Alive);
ADVANCE(T#200ms);
b(PartnerBeat := FALSE, Period := T#1s, Timeout := T#3s);
ASSERT_FALSE(b.Alive);
ASSERT_EQ(UDINT#1, b.LostCount);
b(PartnerBeat := FALSE, Period := T#1s, Timeout := T#3s);
ASSERT_EQ(UDINT#1, b.LostCount);
(* it beats again *)
b(PartnerBeat := TRUE, Period := T#1s, Timeout := T#3s);
ASSERT_TRUE(b.Alive);
END_TEST

TEST heartbeat_from_a_partner_that_starts_high
VAR b : RB_Heartbeat; END_VAR
b(PartnerBeat := TRUE, Period := T#1s, Timeout := T#2s);
ADVANCE(T#1500ms);
b(PartnerBeat := TRUE, Period := T#1s, Timeout := T#2s);
ASSERT_TRUE(b.Alive);
ADVANCE(T#600ms);
b(PartnerBeat := TRUE, Period := T#1s, Timeout := T#2s);
ASSERT_FALSE(b.Alive);
END_TEST

(* ---- ok_rb_light.st ---- *)
(* spec: [blocks.interlock] [blocks.testable]
   expect: ok
   libraries: RootBlocks *)
(* Test suite of RB_Light (F04.LIGHT). Every call passes the inputs that
   matter: block inputs keep their last value. *)
TEST light_toggle_on_off
VAR l : RB_Light; END_VAR
l();
ASSERT_FALSE(l.Out OR l.IsOn);
l(Toggle := TRUE);
ASSERT_TRUE(l.Out AND l.IsOn);
ASSERT_EQ(UDINT#1, l.Switchings);
l(Toggle := FALSE);
ASSERT_TRUE(l.Out);
l(Toggle := TRUE);
ASSERT_FALSE(l.Out);
l(Toggle := FALSE, SetOn := TRUE);
ASSERT_TRUE(l.Out);
ASSERT_EQ(UDINT#2, l.Switchings);
(* off wins over on in the same call *)
l(SetOn := FALSE);
l(SetOn := TRUE, SetOff := TRUE);
ASSERT_FALSE(l.Out);
l(SetOn := FALSE, SetOff := FALSE);
ASSERT_FALSE(l.Out);
(* on while on: no new switch-on *)
l(SetOn := TRUE);
l(SetOn := FALSE);
l(SetOn := TRUE);
ASSERT_EQ(UDINT#3, l.Switchings);
END_TEST

TEST light_stairwell_timer
VAR l : RB_Light; END_VAR
l(SetOn := TRUE, OnTime := T#60s);
ASSERT_EQ(T#60s, l.Remaining);
ADVANCE(T#59s);
l(SetOn := FALSE);
ASSERT_TRUE(l.Out);
ASSERT_EQ(T#1s, l.Remaining);
(* pressing again restarts the time *)
l(SetOn := TRUE);
ASSERT_EQ(T#60s, l.Remaining);
ADVANCE(T#59999ms);
l(SetOn := FALSE);
ASSERT_TRUE(l.Out);
ADVANCE(T#1ms);
l();
ASSERT_FALSE(l.Out OR l.IsOn);
ASSERT_EQ(T#0s, l.Remaining);
(* toggling off a timed light, and on again *)
l(Toggle := TRUE);
ASSERT_TRUE(l.Out);
ADVANCE(T#30s);
l(Toggle := FALSE);
l(Toggle := TRUE);
ASSERT_FALSE(l.Out);
l(Toggle := FALSE);
l(Toggle := TRUE);
ASSERT_EQ(T#60s, l.Remaining);
(* without a time it stays on *)
l(Toggle := FALSE, OnTime := T#0s);
ADVANCE(T#10h);
l();
ASSERT_TRUE(l.Out);
ASSERT_EQ(T#0s, l.Remaining);
END_TEST

TEST light_flash_test_and_interlock
VAR l : RB_Light; END_VAR
l(SetOn := TRUE, Flash := TRUE, FlashTime := T#500ms);
ASSERT_TRUE(l.Out);
ADVANCE(T#500ms);
l();
ASSERT_FALSE(l.Out);
ASSERT_TRUE(l.IsOn);
ADVANCE(T#500ms);
l();
ASSERT_TRUE(l.Out);
l(Flash := FALSE);
ASSERT_TRUE(l.Out);
(* flashing switched on later starts with the lamp on *)
ADVANCE(T#700ms);
l();
l(Flash := TRUE);
ASSERT_TRUE(l.Out);
l(Flash := FALSE);
(* interlock: off now and stays off *)
l(Interlock := TRUE);
ASSERT_FALSE(l.Out OR l.IsOn);
l(Interlock := FALSE);
ASSERT_FALSE(l.Out);
l(SetOn := FALSE);
l(SetOn := TRUE, Interlock := TRUE);
ASSERT_FALSE(l.Out);
(* lamp test lights it whatever the state *)
l(SetOn := FALSE, Interlock := FALSE, LampTest := TRUE);
ASSERT_TRUE(l.Out);
ASSERT_FALSE(l.IsOn);
l(LampTest := FALSE);
ASSERT_FALSE(l.Out);
END_TEST

TEST light_burning_time
VAR l : RB_Light; i : INT; END_VAR
l();
ADVANCE(T#10s);
l(SetOn := TRUE);
ASSERT_TRUE(ABS(l.BurnTime) < 0.001);
ADVANCE(T#2s);
l(SetOn := FALSE);
ASSERT_TRUE(ABS(l.BurnTime - 2.0) < 0.001);
ADVANCE(T#3s);
l(SetOff := TRUE);
ASSERT_TRUE(ABS(l.BurnTime - 5.0) < 0.001);
ADVANCE(T#4s);
l(SetOff := FALSE);
ASSERT_TRUE(ABS(l.BurnTime - 5.0) < 0.001);
(* flashing burns half the time *)
l(SetOn := TRUE, Flash := TRUE, FlashTime := T#1s);
FOR i := 1 TO 4 DO
    ADVANCE(T#1s);
    l(SetOn := FALSE);
END_FOR;
ASSERT_TRUE(ABS(l.BurnTime - 7.0) < 0.001);
END_TEST

(* ---- ok_rb_machine.st ---- *)
(* spec: [blocks.mode] [blocks.command] [blocks.testable]
   expect: ok
   libraries: RootBlocks *)
(* Test suites of RB_ModeManager (F10.MODES), RB_MachineState (F10.STATE)
   and RB_Counter (F03.COUNTER). Every call passes the inputs that matter:
   block inputs keep their last value. *)
TEST modes_requests_and_permissions
VAR m : RB_ModeManager; END_VAR
m();
ASSERT_TRUE(m.Mode = RB_MODE#Off);
ASSERT_FALSE(m.ModeChanged);
m(ReqManual := TRUE);
ASSERT_TRUE(m.Mode = RB_MODE#Manual);
ASSERT_TRUE(m.ModeChanged);
ASSERT_FALSE(m.Rejected);
m(ReqManual := FALSE, ReqAuto := TRUE);
ASSERT_TRUE(m.Mode = RB_MODE#Auto);
m(ReqAuto := FALSE);
ASSERT_FALSE(m.ModeChanged);
m(ReqOff := TRUE);
ASSERT_TRUE(m.Mode = RB_MODE#Off);
(* Auto not allowed: rejected *)
m(ReqOff := FALSE, ReqAuto := TRUE, AutoAllowed := FALSE);
ASSERT_TRUE(m.Rejected);
ASSERT_TRUE(m.Mode = RB_MODE#Off);
m(ReqAuto := FALSE, AutoAllowed := TRUE);
ASSERT_FALSE(m.Rejected);
(* a fault rejects Auto *)
m(ReqAuto := TRUE, Fault := TRUE);
ASSERT_TRUE(m.Rejected);
ASSERT_TRUE(m.Mode = RB_MODE#Off);
(* Manual not allowed *)
m(ReqAuto := FALSE, Fault := FALSE, ReqManual := TRUE, ManualAllowed := FALSE);
ASSERT_TRUE(m.Rejected);
ASSERT_TRUE(m.Mode = RB_MODE#Off);
END_TEST

TEST modes_fall_back_to_off
VAR m : RB_ModeManager; END_VAR
m(ReqAuto := TRUE);
ASSERT_TRUE(m.Mode = RB_MODE#Auto);
m(ReqAuto := FALSE, Fault := TRUE);
ASSERT_TRUE(m.Mode = RB_MODE#Off);
ASSERT_TRUE(m.ModeChanged);
m(Fault := FALSE, ReqAuto := TRUE);
m(ReqAuto := FALSE, AutoAllowed := FALSE);
ASSERT_TRUE(m.Mode = RB_MODE#Off);
m(AutoAllowed := TRUE, ReqManual := TRUE);
ASSERT_TRUE(m.Mode = RB_MODE#Manual);
(* Manual survives a machine fault, but not losing its permission *)
m(ReqManual := FALSE, Fault := TRUE);
ASSERT_TRUE(m.Mode = RB_MODE#Manual);
m(Fault := FALSE, ManualAllowed := FALSE);
ASSERT_TRUE(m.Mode = RB_MODE#Off);
END_TEST

TEST modes_emergency_stop_forces_off
VAR m : RB_ModeManager; END_VAR
m(ReqAuto := TRUE);
m(ReqAuto := FALSE, EStopOk := FALSE);
ASSERT_TRUE(m.Mode = RB_MODE#Off);
m(ReqManual := TRUE, EStopOk := FALSE);
ASSERT_TRUE(m.Rejected);
ASSERT_TRUE(m.Mode = RB_MODE#Off);
m(ReqManual := FALSE, ReqAuto := TRUE, EStopOk := FALSE);
ASSERT_TRUE(m.Rejected);
(* back to normal: the mode stays Off until a new request *)
m(ReqAuto := FALSE, EStopOk := TRUE);
ASSERT_TRUE(m.Mode = RB_MODE#Off);
ASSERT_FALSE(m.Rejected);
m(EStopOk := FALSE);
ASSERT_FALSE(m.Rejected);
END_TEST

TEST machine_state_normal_cycle
VAR s : RB_MachineState; END_VAR
s();
ASSERT_TRUE(s.State = RB_MACHINE_STATE#Stopped);
s(Reset := TRUE);
ASSERT_TRUE(s.State = RB_MACHINE_STATE#Resetting);
s(Reset := FALSE, ResetDone := TRUE);
ASSERT_TRUE(s.State = RB_MACHINE_STATE#Idle);
s(ResetDone := FALSE, Start := TRUE);
ASSERT_TRUE(s.State = RB_MACHINE_STATE#Starting);
ASSERT_FALSE(s.Producing);
s(Start := FALSE, StartDone := TRUE);
ASSERT_TRUE(s.State = RB_MACHINE_STATE#Execute);
ASSERT_TRUE(s.Producing);
s(StartDone := FALSE, Hold := TRUE);
ASSERT_TRUE(s.State = RB_MACHINE_STATE#Held);
s(Hold := FALSE, Unhold := TRUE);
ASSERT_TRUE(s.State = RB_MACHINE_STATE#Execute);
s(Unhold := FALSE, Stop := TRUE);
ASSERT_TRUE(s.State = RB_MACHINE_STATE#Stopping);
s(Stop := FALSE, StopDone := TRUE);
ASSERT_TRUE(s.State = RB_MACHINE_STATE#Stopped);
ASSERT_FALSE(s.Rejected);
END_TEST

TEST machine_state_done_inputs_only_in_their_state
VAR s : RB_MachineState; END_VAR
s(ResetDone := TRUE, StartDone := TRUE, StopDone := TRUE);
ASSERT_TRUE(s.State = RB_MACHINE_STATE#Stopped);
s(ResetDone := FALSE, StartDone := FALSE, StopDone := FALSE, Reset := TRUE);
s(Reset := FALSE, StartDone := TRUE, StopDone := TRUE);
ASSERT_TRUE(s.State = RB_MACHINE_STATE#Resetting);
s(StartDone := FALSE, StopDone := FALSE, ResetDone := TRUE);
s(ResetDone := FALSE, Start := TRUE);
s(Start := FALSE, ResetDone := TRUE, StopDone := TRUE);
ASSERT_TRUE(s.State = RB_MACHINE_STATE#Starting);
s(ResetDone := FALSE, StopDone := FALSE, Stop := TRUE);
ASSERT_TRUE(s.State = RB_MACHINE_STATE#Stopping);
s(Stop := FALSE, ResetDone := TRUE, StartDone := TRUE);
ASSERT_TRUE(s.State = RB_MACHINE_STATE#Stopping);
END_TEST

TEST machine_state_abort_clear_and_rejected
VAR s : RB_MachineState; END_VAR
(* rejected in Stopped *)
s(Start := TRUE);
ASSERT_TRUE(s.Rejected);
s(Start := FALSE, Stop := TRUE);
ASSERT_TRUE(s.Rejected);
s(Stop := FALSE, Hold := TRUE);
ASSERT_TRUE(s.Rejected);
s(Hold := FALSE, Unhold := TRUE);
ASSERT_TRUE(s.Rejected);
s(Unhold := FALSE, Clear := TRUE);
ASSERT_TRUE(s.Rejected);
s(Clear := FALSE);
ASSERT_FALSE(s.Rejected);
(* abort from any state, clear back to Stopped *)
s(Abort := TRUE);
ASSERT_TRUE(s.State = RB_MACHINE_STATE#Aborted);
s(Abort := FALSE);
s(Abort := TRUE);
ASSERT_TRUE(s.Rejected);
s(Abort := FALSE, Reset := TRUE);
ASSERT_TRUE(s.Rejected);
s(Reset := FALSE, Clear := TRUE);
ASSERT_TRUE(s.State = RB_MACHINE_STATE#Stopped);
(* stop from Idle, Starting and Held *)
s(Clear := FALSE, Reset := TRUE);
s(Reset := FALSE, ResetDone := TRUE);
s(ResetDone := FALSE, Stop := TRUE);
ASSERT_TRUE(s.State = RB_MACHINE_STATE#Stopping);
s(Stop := FALSE, StopDone := TRUE);
s(StopDone := FALSE, Reset := TRUE);
ASSERT_TRUE(s.State = RB_MACHINE_STATE#Resetting);
s(Reset := FALSE);
s(Reset := TRUE);
ASSERT_TRUE(s.Rejected);
s(Reset := FALSE, ResetDone := TRUE);
s(ResetDone := FALSE, Start := TRUE);
s(Start := FALSE, Stop := TRUE);
ASSERT_TRUE(s.State = RB_MACHINE_STATE#Stopping);
s(Stop := FALSE, StopDone := TRUE);
s(StopDone := FALSE, Reset := TRUE);
s(Reset := FALSE, ResetDone := TRUE);
s(ResetDone := FALSE, Start := TRUE);
s(Start := FALSE, StartDone := TRUE);
s(StartDone := FALSE, Hold := TRUE);
s(Hold := FALSE, Stop := TRUE);
ASSERT_TRUE(s.State = RB_MACHINE_STATE#Stopping);
s(Stop := FALSE, Hold := TRUE);
ASSERT_TRUE(s.Rejected);
s(Hold := FALSE, Abort := TRUE);
ASSERT_TRUE(s.State = RB_MACHINE_STATE#Aborted);
END_TEST

TEST counter_counts_to_preset
VAR c : RB_Counter; END_VAR
c(In := FALSE, Preset := 3);
ASSERT_EQ(UDINT#3, c.Remaining);
c(In := TRUE, Preset := 3);
c(In := TRUE, Preset := 3);
ASSERT_EQ(UDINT#1, c.Count);
c(In := FALSE, Preset := 3);
c(In := TRUE, Preset := 3);
ASSERT_EQ(UDINT#2, c.Count);
ASSERT_FALSE(c.Done);
ASSERT_EQ(UDINT#1, c.Remaining);
c(In := FALSE, Preset := 3);
c(In := TRUE, Preset := 3);
ASSERT_TRUE(c.Done);
ASSERT_TRUE(c.BatchDone);
ASSERT_EQ(UDINT#1, c.Batches);
ASSERT_EQ(UDINT#0, c.Remaining);
c(In := FALSE, Preset := 3);
ASSERT_FALSE(c.BatchDone);
(* without auto restart it stays at the preset; the total goes on *)
c(In := TRUE, Preset := 3);
ASSERT_EQ(UDINT#3, c.Count);
ASSERT_EQ(UDINT#4, c.Total);
ASSERT_EQ(UDINT#1, c.Batches);
c(In := FALSE, Preset := 3, Reset := TRUE);
ASSERT_EQ(UDINT#0, c.Count);
ASSERT_FALSE(c.Done);
ASSERT_EQ(UDINT#4, c.Total);
END_TEST

TEST counter_batches_with_auto_restart
VAR c : RB_Counter; i : INT; END_VAR
FOR i := 1 TO 7 DO
    c(In := TRUE, Preset := 2, AutoRestart := TRUE);
    c(In := FALSE, Preset := 2, AutoRestart := TRUE);
END_FOR;
ASSERT_EQ(UDINT#3, c.Batches);
ASSERT_EQ(UDINT#1, c.Count);
ASSERT_EQ(UDINT#7, c.Total);
c(In := TRUE, Preset := 2, AutoRestart := TRUE);
ASSERT_TRUE(c.BatchDone);
ASSERT_TRUE(c.Done);
ASSERT_EQ(UDINT#4, c.Batches);
(* a preset lowered below the count: done at once *)
c(In := FALSE, Preset := 1, AutoRestart := FALSE, Reset := FALSE);
ASSERT_TRUE(c.Done);
ASSERT_EQ(UDINT#0, c.Remaining);
END_TEST

(* ---- ok_rb_motor.st ---- *)
(* spec: [blocks.command] [blocks.mode] [blocks.interlock] [blocks.fault] [blocks.feedback] [blocks.status]
   expect: ok
   libraries: RootBlocks *)
(* Test suite of RB_Motor (card blocks/cards/F04.MOTOR.DOL.md). Every call
   passes the inputs that matter: block inputs keep their last value. *)
TEST motor_starts_and_reports
VAR m : RB_Motor; END_VAR
m(Mode := RB_MODE#Auto, AutoRun := TRUE, FbRunning := FALSE);
ASSERT_TRUE(m.Run);
ASSERT_FALSE(m.Running);
ASSERT_TRUE(m.Status.Commanded);
m(Mode := RB_MODE#Auto, AutoRun := TRUE, FbRunning := TRUE);
ASSERT_TRUE(m.Running);
ASSERT_TRUE(m.Status.Active);
ASSERT_EQ(UDINT#1, m.Status.Starts);
ASSERT_TRUE(m.Status.Mode = RB_MODE#Auto);
m(Mode := RB_MODE#Auto, AutoRun := FALSE, FbRunning := TRUE);
ASSERT_FALSE(m.Run);
m(Mode := RB_MODE#Auto, AutoRun := FALSE, FbRunning := FALSE);
m(Mode := RB_MODE#Auto, AutoRun := TRUE, FbRunning := FALSE);
ASSERT_EQ(UDINT#2, m.Status.Starts);
ASSERT_FALSE(m.Error);
ASSERT_FALSE(m.Status.Error);
END_TEST

TEST motor_mode_interlock_permissive
VAR m : RB_Motor; END_VAR
m(Mode := RB_MODE#Auto, ManRun := TRUE, FbRunning := FALSE);
ASSERT_FALSE(m.Run);
m(Mode := RB_MODE#Manual, ManRun := TRUE, AutoRun := FALSE, FbRunning := FALSE);
ASSERT_TRUE(m.Run);
m(Mode := RB_MODE#Manual, ManRun := TRUE, Interlock := TRUE, FbRunning := TRUE);
ASSERT_FALSE(m.Run);
m(Mode := RB_MODE#Off, ManRun := TRUE, AutoRun := TRUE, Interlock := FALSE, FbRunning := FALSE);
ASSERT_FALSE(m.Run);
m(Mode := RB_MODE#Auto, AutoRun := TRUE, Permissive := FALSE, FbRunning := FALSE);
ASSERT_FALSE(m.Run);
m(Mode := RB_MODE#Auto, AutoRun := TRUE, Permissive := TRUE, FbRunning := FALSE);
ASSERT_TRUE(m.Run);
m(Mode := RB_MODE#Auto, AutoRun := TRUE, Permissive := FALSE, FbRunning := TRUE);
ASSERT_TRUE(m.Run);
END_TEST

TEST motor_overload_trips_at_once_and_latches
VAR m : RB_Motor; END_VAR
m(Mode := RB_MODE#Auto, AutoRun := TRUE, FbRunning := TRUE);
m(Mode := RB_MODE#Auto, AutoRun := TRUE, FbRunning := TRUE, Overload := TRUE);
ASSERT_FALSE(m.Run);
ASSERT_TRUE(m.Error);
ASSERT_EQ(UDINT#3, m.ErrorID);
m(Mode := RB_MODE#Auto, AutoRun := TRUE, FbRunning := FALSE, Overload := FALSE);
ASSERT_TRUE(m.Error);
ASSERT_FALSE(m.Run);
(* reset while still tripped: the fault returns at once *)
m(Mode := RB_MODE#Auto, AutoRun := TRUE, FbRunning := FALSE, Overload := TRUE, Reset := TRUE);
ASSERT_TRUE(m.Error);
m(Mode := RB_MODE#Auto, AutoRun := TRUE, FbRunning := FALSE, Overload := FALSE, Reset := FALSE);
m(Mode := RB_MODE#Auto, AutoRun := TRUE, FbRunning := FALSE, Overload := FALSE, Reset := TRUE);
ASSERT_FALSE(m.Error);
ASSERT_EQ(UDINT#0, m.ErrorID);
ASSERT_TRUE(m.Run);
END_TEST

TEST motor_no_running_feedback
VAR m : RB_Motor; END_VAR
m(Mode := RB_MODE#Auto, AutoRun := TRUE, FbRunning := FALSE, FeedbackTime := T#1s);
ADVANCE(T#900ms);
m(Mode := RB_MODE#Auto, AutoRun := TRUE, FbRunning := FALSE, FeedbackTime := T#1s);
ASSERT_FALSE(m.Error);
ADVANCE(T#200ms);
m(Mode := RB_MODE#Auto, AutoRun := TRUE, FbRunning := FALSE, FeedbackTime := T#1s);
ASSERT_TRUE(m.Error);
ASSERT_EQ(UDINT#1, m.ErrorID);
ASSERT_FALSE(m.Run);
ASSERT_EQ(UDINT#1, m.Status.ErrorID);
END_TEST

TEST motor_contactor_stuck
VAR m : RB_Motor; END_VAR
m(Mode := RB_MODE#Auto, AutoRun := FALSE, FbRunning := TRUE, FeedbackTime := T#1s);
ADVANCE(T#1100ms);
m(Mode := RB_MODE#Auto, AutoRun := FALSE, FbRunning := TRUE, FeedbackTime := T#1s);
ASSERT_TRUE(m.Error);
ASSERT_EQ(UDINT#2, m.ErrorID);
END_TEST

TEST motor_restart_delay
VAR m : RB_Motor; END_VAR
m(Mode := RB_MODE#Auto, AutoRun := FALSE, FbRunning := FALSE, RestartDelay := T#10s);
ADVANCE(T#11s);
m(Mode := RB_MODE#Auto, AutoRun := TRUE, FbRunning := FALSE, RestartDelay := T#10s);
ASSERT_TRUE(m.Run);
m(Mode := RB_MODE#Auto, AutoRun := FALSE, FbRunning := TRUE, RestartDelay := T#10s);
ADVANCE(T#5s);
m(Mode := RB_MODE#Auto, AutoRun := TRUE, FbRunning := FALSE, RestartDelay := T#10s);
ASSERT_FALSE(m.Run);
ASSERT_EQ(UDINT#1, m.Status.Starts);
ADVANCE(T#6s);
m(Mode := RB_MODE#Auto, AutoRun := TRUE, FbRunning := FALSE, RestartDelay := T#10s);
ASSERT_TRUE(m.Run);
ASSERT_EQ(UDINT#2, m.Status.Starts);
END_TEST

TEST motor_without_feedback
VAR m : RB_Motor; END_VAR
m(Mode := RB_MODE#Auto, AutoRun := TRUE, Feedback := FALSE, FbRunning := FALSE, FeedbackTime := T#1s);
ASSERT_TRUE(m.Running);
ADVANCE(T#5s);
m(Mode := RB_MODE#Auto, AutoRun := TRUE, Feedback := FALSE, FbRunning := FALSE, FeedbackTime := T#1s);
ASSERT_FALSE(m.Error);
(* switching supervision on starts its timer fresh *)
m(Mode := RB_MODE#Auto, AutoRun := TRUE, Feedback := TRUE, FbRunning := FALSE, FeedbackTime := T#1s);
ASSERT_FALSE(m.Error);
ASSERT_FALSE(m.Running);
END_TEST

TEST motor_runs_normally_past_the_feedback_time
VAR m : RB_Motor; END_VAR
m(Mode := RB_MODE#Auto, AutoRun := TRUE, FbRunning := TRUE, FeedbackTime := T#1s);
ADVANCE(T#3s);
m(Mode := RB_MODE#Auto, AutoRun := TRUE, FbRunning := TRUE, FeedbackTime := T#1s);
ASSERT_FALSE(m.Error);
ASSERT_TRUE(m.Run);
END_TEST

(* ---- ok_rb_motor_reversing.st ---- *)
(* spec: [blocks.command] [blocks.mode] [blocks.interlock] [blocks.fault] [blocks.feedback] [blocks.status]
   expect: ok
   libraries: RootBlocks *)
(* Test suite of RB_MotorReversing (card blocks/cards/F04.MOTOR.REV.md).
   Every call passes the inputs that matter: block inputs keep their last
   value. *)
TEST reversing_forward_then_reverse_with_dead_time
VAR m : RB_MotorReversing; i : INT; both : BOOL; END_VAR
m(Mode := RB_MODE#Auto, AutoFwd := TRUE, AutoRev := FALSE, FbFwd := FALSE, FbRev := FALSE, ReverseDelay := T#1s);
ASSERT_FALSE(m.RunFwd);
ADVANCE(T#1s);
m(Mode := RB_MODE#Auto, AutoFwd := TRUE, AutoRev := FALSE, FbFwd := FALSE, FbRev := FALSE, ReverseDelay := T#1s);
ASSERT_TRUE(m.RunFwd);
ASSERT_TRUE(m.Status.Commanded);
m(Mode := RB_MODE#Auto, AutoFwd := TRUE, AutoRev := FALSE, FbFwd := TRUE, FbRev := FALSE, ReverseDelay := T#1s);
ASSERT_TRUE(m.RunningFwd);
ASSERT_FALSE(m.RunningRev);
ASSERT_TRUE(m.Status.Active);
ASSERT_EQ(UDINT#1, m.Status.Starts);
(* reverse: forward drops at once, reverse waits for the dead time *)
m(Mode := RB_MODE#Auto, AutoFwd := FALSE, AutoRev := TRUE, FbFwd := TRUE, FbRev := FALSE, ReverseDelay := T#1s);
ASSERT_FALSE(m.RunFwd);
ASSERT_FALSE(m.RunRev);
FOR i := 1 TO 9 DO
    ADVANCE(T#100ms);
    m(Mode := RB_MODE#Auto, AutoFwd := FALSE, AutoRev := TRUE, FbFwd := FALSE, FbRev := FALSE, ReverseDelay := T#1s);
    IF m.RunRev THEN both := TRUE; END_IF;
END_FOR;
ASSERT_FALSE(both);
ADVANCE(T#200ms);
m(Mode := RB_MODE#Auto, AutoFwd := FALSE, AutoRev := TRUE, FbFwd := FALSE, FbRev := FALSE, ReverseDelay := T#1s);
ASSERT_TRUE(m.RunRev);
ASSERT_FALSE(m.RunFwd);
ASSERT_EQ(UDINT#2, m.Status.Starts);
m(Mode := RB_MODE#Auto, AutoFwd := FALSE, AutoRev := TRUE, FbFwd := FALSE, FbRev := TRUE, ReverseDelay := T#1s);
ASSERT_TRUE(m.RunningRev);
ASSERT_FALSE(m.Error);
END_TEST

TEST reversing_both_commands_stop
VAR m : RB_MotorReversing; END_VAR
m(Mode := RB_MODE#Auto, AutoFwd := TRUE, AutoRev := FALSE, ReverseDelay := T#0s);
ASSERT_TRUE(m.RunFwd);
m(Mode := RB_MODE#Auto, AutoFwd := TRUE, AutoRev := TRUE, FbFwd := TRUE, ReverseDelay := T#0s);
ASSERT_FALSE(m.RunFwd);
ASSERT_FALSE(m.RunRev);
END_TEST

TEST reversing_modes_interlock_permissive
VAR m : RB_MotorReversing; END_VAR
m(Mode := RB_MODE#Auto, ManRev := TRUE, ReverseDelay := T#0s);
ASSERT_FALSE(m.RunRev);
m(Mode := RB_MODE#Manual, ManRev := TRUE, ManFwd := FALSE, ReverseDelay := T#0s);
ASSERT_TRUE(m.RunRev);
m(Mode := RB_MODE#Manual, ManRev := TRUE, Interlock := TRUE, FbRev := TRUE, ReverseDelay := T#0s);
ASSERT_FALSE(m.RunRev);
m(Mode := RB_MODE#Manual, ManFwd := TRUE, ManRev := FALSE, Interlock := FALSE, FbRev := FALSE, ReverseDelay := T#0s);
ASSERT_TRUE(m.RunFwd);
m(Mode := RB_MODE#Off, ManFwd := TRUE, FbFwd := TRUE, ReverseDelay := T#0s);
ASSERT_FALSE(m.RunFwd);
m(Mode := RB_MODE#Auto, AutoRev := TRUE, Permissive := FALSE, FbFwd := FALSE, ReverseDelay := T#0s);
ASSERT_FALSE(m.RunRev);
m(Mode := RB_MODE#Auto, AutoFwd := TRUE, AutoRev := FALSE, Permissive := FALSE, ReverseDelay := T#0s);
ASSERT_FALSE(m.RunFwd);
m(Mode := RB_MODE#Auto, AutoFwd := TRUE, Permissive := TRUE, ReverseDelay := T#0s);
ASSERT_TRUE(m.RunFwd);
m(Mode := RB_MODE#Auto, AutoFwd := TRUE, Permissive := FALSE, FbFwd := TRUE, ReverseDelay := T#0s);
ASSERT_TRUE(m.RunFwd);
m(Mode := RB_MODE#Auto, AutoFwd := FALSE, AutoRev := TRUE, Permissive := TRUE, FbFwd := FALSE, ReverseDelay := T#0s);
m(Mode := RB_MODE#Auto, AutoFwd := FALSE, AutoRev := TRUE, Permissive := TRUE, FbFwd := FALSE, ReverseDelay := T#0s);
ASSERT_TRUE(m.RunRev);
m(Mode := RB_MODE#Auto, AutoRev := TRUE, Permissive := FALSE, FbRev := TRUE, ReverseDelay := T#0s);
ASSERT_TRUE(m.RunRev);
END_TEST

TEST reversing_faults
VAR m : RB_MotorReversing; n : RB_MotorReversing; k : RB_MotorReversing; o : RB_MotorReversing; END_VAR
(* no feedback for the commanded direction *)
m(Mode := RB_MODE#Auto, AutoRev := TRUE, FbRev := FALSE, ReverseDelay := T#0s, FeedbackTime := T#1s);
ADVANCE(T#1100ms);
m(Mode := RB_MODE#Auto, AutoRev := TRUE, FbRev := FALSE, ReverseDelay := T#0s, FeedbackTime := T#1s);
ASSERT_TRUE(m.Error);
ASSERT_EQ(UDINT#1, m.ErrorID);
ASSERT_FALSE(m.RunRev);
ASSERT_EQ(UDINT#1, m.Status.ErrorID);
ASSERT_TRUE(m.Status.Error);
(* forward feedback without a command *)
n(Mode := RB_MODE#Auto, FbFwd := TRUE, ReverseDelay := T#0s, FeedbackTime := T#1s);
ADVANCE(T#1100ms);
n(Mode := RB_MODE#Auto, FbFwd := TRUE, ReverseDelay := T#0s, FeedbackTime := T#1s);
ASSERT_EQ(UDINT#2, n.ErrorID);
ASSERT_TRUE(n.Error);
(* both feedback contacts *)
k(Mode := RB_MODE#Auto, AutoFwd := TRUE, FbFwd := TRUE, FbRev := TRUE, ReverseDelay := T#0s, FeedbackTime := T#1s);
ASSERT_FALSE(k.RunningFwd);
ASSERT_FALSE(k.RunningRev);
ADVANCE(T#1100ms);
k(Mode := RB_MODE#Auto, AutoFwd := TRUE, FbFwd := TRUE, FbRev := TRUE, ReverseDelay := T#0s, FeedbackTime := T#1s);
ASSERT_EQ(UDINT#4, k.ErrorID);
ASSERT_FALSE(k.RunFwd);
(* overload, then reset *)
o(Mode := RB_MODE#Auto, AutoFwd := TRUE, Overload := TRUE, ReverseDelay := T#0s);
ASSERT_EQ(UDINT#3, o.ErrorID);
ASSERT_FALSE(o.RunFwd);
o(Mode := RB_MODE#Auto, AutoFwd := TRUE, Overload := FALSE, Reset := TRUE, ReverseDelay := T#0s);
ASSERT_FALSE(o.Error);
ASSERT_EQ(UDINT#0, o.ErrorID);
ASSERT_TRUE(o.RunFwd);
END_TEST

TEST reversing_without_feedback
VAR m : RB_MotorReversing; END_VAR
m(Mode := RB_MODE#Auto, AutoFwd := TRUE, Feedback := FALSE, ReverseDelay := T#0s, FeedbackTime := T#1s);
ASSERT_TRUE(m.RunningFwd);
ADVANCE(T#5s);
m(Mode := RB_MODE#Auto, AutoFwd := FALSE, AutoRev := TRUE, Feedback := FALSE, ReverseDelay := T#0s, FeedbackTime := T#1s);
m(Mode := RB_MODE#Auto, AutoFwd := FALSE, AutoRev := TRUE, Feedback := FALSE, ReverseDelay := T#0s, FeedbackTime := T#1s);
ASSERT_TRUE(m.RunningRev);
ASSERT_FALSE(m.Error);
m(Mode := RB_MODE#Auto, AutoRev := TRUE, Feedback := TRUE, FbRev := FALSE, ReverseDelay := T#0s, FeedbackTime := T#1s);
ASSERT_FALSE(m.Error);
END_TEST

TEST reversing_details
VAR m : RB_MotorReversing; s : RB_MotorReversing; o : RB_MotorReversing; END_VAR
(* both commands from standstill: nothing runs *)
s(Mode := RB_MODE#Auto, AutoFwd := TRUE, AutoRev := TRUE, ReverseDelay := T#0s);
ASSERT_FALSE(s.RunFwd);
ASSERT_FALSE(s.RunRev);
(* Off: no direction runs *)
o(Mode := RB_MODE#Off, ManRev := TRUE, AutoRev := TRUE, ReverseDelay := T#0s);
ASSERT_FALSE(o.RunRev);
(* forward runs normally past the feedback time; starts counted once *)
m(Mode := RB_MODE#Auto, AutoFwd := TRUE, FbFwd := TRUE, ReverseDelay := T#0s, FeedbackTime := T#1s);
m(Mode := RB_MODE#Auto, AutoFwd := TRUE, FbFwd := TRUE, ReverseDelay := T#0s, FeedbackTime := T#1s);
ADVANCE(T#3s);
m(Mode := RB_MODE#Auto, AutoFwd := TRUE, FbFwd := TRUE, ReverseDelay := T#0s, FeedbackTime := T#1s);
ASSERT_FALSE(m.Error);
ASSERT_EQ(UDINT#1, m.Status.Starts);
(* an interlock stops forward too *)
m(Mode := RB_MODE#Auto, AutoFwd := TRUE, FbFwd := TRUE, Interlock := TRUE, ReverseDelay := T#0s, FeedbackTime := T#1s);
ASSERT_FALSE(m.RunFwd);
m(Mode := RB_MODE#Auto, AutoFwd := FALSE, FbFwd := FALSE, Interlock := FALSE, ReverseDelay := T#0s, FeedbackTime := T#1s);
(* reverse runs normally past the feedback time *)
m(Mode := RB_MODE#Auto, AutoRev := TRUE, FbRev := TRUE, ReverseDelay := T#0s, FeedbackTime := T#1s);
ADVANCE(T#3s);
m(Mode := RB_MODE#Auto, AutoRev := TRUE, FbRev := TRUE, ReverseDelay := T#0s, FeedbackTime := T#1s);
ASSERT_FALSE(m.Error);
ASSERT_TRUE(m.RunRev);
END_TEST

TEST reversing_supervision_switched_on_starts_fresh
VAR m : RB_MotorReversing; k : RB_MotorReversing; END_VAR
m(Mode := RB_MODE#Auto, AutoFwd := TRUE, Feedback := FALSE, FbFwd := FALSE, ReverseDelay := T#0s, FeedbackTime := T#1s);
ADVANCE(T#5s);
m(Mode := RB_MODE#Auto, AutoFwd := TRUE, Feedback := FALSE, FbFwd := FALSE, ReverseDelay := T#0s, FeedbackTime := T#1s);
m(Mode := RB_MODE#Auto, AutoFwd := TRUE, Feedback := TRUE, FbFwd := FALSE, ReverseDelay := T#0s, FeedbackTime := T#1s);
ASSERT_FALSE(m.Error);
k(Mode := RB_MODE#Auto, AutoFwd := TRUE, Feedback := FALSE, FbFwd := TRUE, FbRev := TRUE, ReverseDelay := T#0s, FeedbackTime := T#1s);
ADVANCE(T#5s);
k(Mode := RB_MODE#Auto, AutoFwd := TRUE, Feedback := FALSE, FbFwd := TRUE, FbRev := TRUE, ReverseDelay := T#0s, FeedbackTime := T#1s);
k(Mode := RB_MODE#Auto, AutoFwd := TRUE, Feedback := TRUE, FbFwd := TRUE, FbRev := TRUE, ReverseDelay := T#0s, FeedbackTime := T#1s);
ASSERT_FALSE(k.Error);
ADVANCE(T#1100ms);
k(Mode := RB_MODE#Auto, AutoFwd := TRUE, Feedback := TRUE, FbFwd := TRUE, FbRev := TRUE, ReverseDelay := T#0s, FeedbackTime := T#1s);
ASSERT_TRUE(k.Error);
ASSERT_EQ(UDINT#4, k.ErrorID);
END_TEST
